--- program plaizgr (robot Fanuc LR Mate 200iD/7L) ---
  Suave(1)
  Establecer velocidad (1000.0 mm/s)
  Est. Ref.: RobotiQ 2F-140 Gripper (Mechanism) Base
  Est. herr: Tool 1
  Mostrar Tool 1
  MoveJ 1 to (362.78, 154.32, 254.42) mm, rotated rx 150.39 ry -54.39 rz -78.94 deg; joints [58.46, 52.97, -15.965, -58.774, -88.343, 127.064]
  MoveL 2 to (362.78, 154.32, 254.42) mm, rotated rx 150.39 ry -54.39 rz -78.94 deg; joints [58.46, 52.97, -15.965, -58.774, -88.343, 127.064]
  MoveL 3 to (343.17, 154.32, 156.36) mm, rotated rx 150.39 ry -54.39 rz -78.94 deg; joints [59.167, 60.189, -23.258, -59.407, -84.021, 132.99]
  MoveL 4 to (343.17, 154.32, 156.36) mm, rotated rx 150.39 ry -54.39 rz -78.94 deg; joints [59.167, 60.189, -23.258, -59.407, -84.021, 132.99]
  Establecer velocidad (50.0 mm/s)
  MoveL 5 to (357.24, 155.51, 156.36) mm, rotated rx 150.39 ry -54.39 rz -78.94 deg; joints [58.593, 58.357, -25.001, -59.364, -83.585, 134.768]
  MoveL 6 to (371.41, 155.49, 156.36) mm, rotated rx 150.39 ry -54.39 rz -78.94 deg; joints [58.07, 56.537, -26.718, -59.336, -83.115, 136.496]
  MoveL 7 to (385.52, 154.28, 156.36) mm, rotated rx 150.39 ry -54.39 rz -78.94 deg; joints [57.607, 54.737, -28.4, -59.33, -82.61, 138.165]
  MoveL 8 to (399.43, 151.88, 156.36) mm, rotated rx 150.39 ry -54.39 rz -78.94 deg; joints [57.21, 52.967, -30.039, -59.349, -82.072, 139.766]
  MoveL 9 to (413.04, 148.32, 157.01) mm, rotated rx 150.39 ry -54.39 rz -78.94 deg; joints [56.883, 51.186, -31.573, -59.393, -81.532, 141.244]
  MoveL 10 to (427.09, 143.6, 159.01) mm, rotated rx 150.39 ry -54.39 rz -78.94 deg; joints [56.601, 49.261, -33.008, -59.45, -81.007, 142.617]
  MoveL 11 to (441.01, 139.44, 162.37) mm, rotated rx 150.39 ry -54.39 rz -78.94 deg; joints [56.277, 47.356, -34.183, -59.457, -80.642, 143.78]
  MoveL 12 to (454.79, 136.05, 167.07) mm, rotated rx 150.39 ry -54.39 rz -78.94 deg; joints [55.897, 45.467, -35.092, -59.397, -80.449, 144.736]
  MoveL 13 to (468.79, 133.33, 171.26) mm, rotated rx 150.39 ry -54.39 rz -78.94 deg; joints [55.448, 43.671, -35.961, -59.295, -80.321, 145.682]
  MoveL 14 to (483.13, 131.27, 174.06) mm, rotated rx 150.39 ry -54.39 rz -78.94 deg; joints [54.922, 42.013, -36.897, -59.158, -80.205, 146.718]
  MoveL 15 to (497.82, 129.91, 175.45) mm, rotated rx 150.39 ry -54.39 rz -78.94 deg; joints [54.312, 40.498, -37.91, -58.981, -80.1, 147.853]
  MoveL 16 to (513.8, 129.29, 175.6) mm, rotated rx 150.39 ry -54.39 rz -78.94 deg; joints [53.565, 39.04, -39.056, -58.741, -80.008, 149.156]
  MoveL 17 to (529.8, 129.54, 175.6) mm, rotated rx 150.39 ry -54.39 rz -78.94 deg; joints [52.727, 37.685, -40.126, -58.427, -80.002, 150.425]
  MoveL 18 to (545.79, 129.54, 175.6) mm, rotated rx 150.39 ry -54.39 rz -78.94 deg; joints [51.873, 36.349, -41.162, -58.086, -80.008, 151.666]
  MoveL 19 to (561.78, 129.54, 175.6) mm, rotated rx 150.39 ry -54.39 rz -78.94 deg; joints [50.985, 35.046, -42.154, -57.706, -80.042, 152.877]
  MoveL 20 to (577.78, 129.54, 175.6) mm, rotated rx 150.39 ry -54.39 rz -78.94 deg; joints [50.063, 33.774, -43.105, -57.286, -80.104, 154.061]
  MoveL 21 to (587.78, 129.54, 175.6) mm, rotated rx 150.39 ry -54.39 rz -78.94 deg; joints [49.468, 32.995, -43.678, -57.001, -80.156, 154.788]
  MoveL 22 to (597.77, 129.54, 175.6) mm, rotated rx 150.39 ry -54.39 rz -78.94 deg; joints [48.857, 32.226, -44.236, -56.7, -80.219, 155.506]
  MoveL 23 to (607.77, 129.54, 175.6) mm, rotated rx 150.39 ry -54.39 rz -78.94 deg; joints [48.232, 31.469, -44.779, -56.382, -80.292, 156.215]
  MoveL 24 to (617.86, 129.25, 175.6) mm, rotated rx 150.39 ry -54.39 rz -78.94 deg; joints [47.606, 30.696, -45.325, -56.058, -80.356, 156.925]
  MoveL 25 to (624.85, 127.52, 175.6) mm, rotated rx 150.39 ry -54.39 rz -78.94 deg; joints [47.271, 30.062, -45.767, -55.904, -80.303, 157.429]
  MoveL 26 to (631.59, 124.12, 175.6) mm, rotated rx 150.39 ry -54.39 rz -78.94 deg; joints [47.066, 29.337, -46.266, -55.841, -80.141, 157.929]
  MoveL 27 to (637.51, 119.15, 175.6) mm, rotated rx 150.39 ry -54.39 rz -78.94 deg; joints [47.027, 28.568, -46.786, -55.891, -79.871, 158.382]
  MoveL 28 to (642.09, 112.97, 175.6) mm, rotated rx 150.39 ry -54.39 rz -78.94 deg; joints [47.169, 27.817, -47.287, -56.061, -79.51, 158.749]
  MoveL 29 to (645.05, 106.13, 175.6) mm, rotated rx 150.39 ry -54.39 rz -78.94 deg; joints [47.477, 27.141, -47.73, -56.336, -79.091, 159.006]
  MoveL 30 to (646.36, 99.2, 175.6) mm, rotated rx 150.39 ry -54.39 rz -78.94 deg; joints [47.914, 26.584, -48.09, -56.687, -78.648, 159.147]
  MoveL 31 to (646.47, 92.51, 175.6) mm, rotated rx 150.39 ry -54.39 rz -78.94 deg; joints [48.424, 26.135, -48.377, -57.079, -78.207, 159.203]
  MoveL 32 to (646.47, 85.85, 175.6) mm, rotated rx 150.39 ry -54.39 rz -78.94 deg; joints [48.949, 25.7, -48.651, -57.481, -77.766, 159.247]
  MoveL 33 to (645.82, 79.04, 175.6) mm, rotated rx 150.39 ry -54.39 rz -78.94 deg; joints [49.539, 25.31, -48.895, -57.924, -77.307, 159.245]
  MoveL 34 to (643.6, 72.09, 175.6) mm, rotated rx 150.39 ry -54.39 rz -78.94 deg; joints [50.256, 25.036, -49.065, -58.442, -76.818, 159.139]
  MoveL 35 to (639.71, 65.55, 175.6) mm, rotated rx 150.39 ry -54.39 rz -78.94 deg; joints [51.058, 24.923, -49.134, -58.997, -76.332, 158.919]
  MoveL 36 to (634.33, 59.99, 175.6) mm, rotated rx 150.39 ry -54.39 rz -78.94 deg; joints [51.88, 24.997, -49.089, -59.541, -75.893, 158.595]
  MoveL 37 to (627.87, 55.87, 175.6) mm, rotated rx 150.39 ry -54.39 rz -78.94 deg; joints [52.646, 25.253, -48.931, -60.02, -75.539, 158.193]
  MoveL 38 to (620.92, 53.42, 175.6) mm, rotated rx 150.39 ry -54.39 rz -78.94 deg; joints [53.296, 25.655, -48.679, -60.397, -75.292, 157.748]
  MoveL 39 to (611.8, 52.57, 175.6) mm, rotated rx 150.39 ry -54.39 rz -78.94 deg; joints [53.933, 26.331, -48.252, -60.721, -75.134, 157.149]
  MoveL 40 to (602.92, 52.57, 175.6) mm, rotated rx 150.39 ry -54.39 rz -78.94 deg; joints [54.47, 27.044, -47.793, -60.966, -75.045, 156.553]
  MoveL 41 to (594.03, 52.57, 175.6) mm, rotated rx 150.39 ry -54.39 rz -78.94 deg; joints [54.993, 27.763, -47.322, -61.196, -74.963, 155.949]
  MoveL 42 to (585.15, 52.57, 175.6) mm, rotated rx 150.39 ry -54.39 rz -78.94 deg; joints [55.503, 28.488, -46.839, -61.411, -74.89, 155.338]
  MoveL 43 to (576.26, 52.57, 175.6) mm, rotated rx 150.39 ry -54.39 rz -78.94 deg; joints [56, 29.22, -46.345, -61.61, -74.826, 154.719]
  MoveL 44 to (567.37, 52.57, 175.6) mm, rotated rx 150.39 ry -54.39 rz -78.94 deg; joints [56.485, 29.958, -45.838, -61.795, -74.77, 154.092]
  MoveL 45 to (549.78, 52.57, 175.6) mm, rotated rx 150.39 ry -54.39 rz -78.94 deg; joints [57.409, 31.439, -44.799, -62.118, -74.685, 152.825]
  MoveL 46 to (532.19, 52.57, 175.6) mm, rotated rx 150.39 ry -54.39 rz -78.94 deg; joints [58.288, 32.948, -43.711, -62.387, -74.634, 151.522]
  MoveL 47 to (514.6, 51.98, 175.6) mm, rotated rx 150.39 ry -54.39 rz -78.94 deg; joints [59.172, 34.456, -42.597, -62.638, -74.577, 150.188]
  MoveL 48 to (497.1, 50.19, 175.42) mm, rotated rx 150.39 ry -54.39 rz -78.94 deg; joints [60.103, 35.943, -41.504, -62.905, -74.462, 148.851]
  MoveL 49 to (482.53, 47.78, 173.97) mm, rotated rx 150.39 ry -54.39 rz -78.94 deg; joints [60.918, 37.26, -40.73, -63.17, -74.265, 147.846]
  MoveL 50 to (468.32, 44.58, 171.14) mm, rotated rx 150.39 ry -54.39 rz -78.94 deg; joints [61.75, 38.633, -40.118, -63.472, -73.975, 146.983]
  MoveL 51 to (454.47, 40.81, 166.96) mm, rotated rx 150.39 ry -54.39 rz -78.94 deg; joints [62.583, 40.068, -39.653, -63.803, -73.608, 146.252]
  MoveL 52 to (440.68, 37.6, 162.27) mm, rotated rx 150.39 ry -54.39 rz -78.94 deg; joints [63.348, 41.583, -39.17, -64.082, -73.29, 145.529]
  MoveL 53 to (426.53, 35.07, 158.91) mm, rotated rx 150.39 ry -54.39 rz -78.94 deg; joints [64.051, 43.092, -38.442, -64.253, -73.114, 144.595]
  MoveL 54 to (412.03, 33.26, 156.92) mm, rotated rx 150.39 ry -54.39 rz -78.94 deg; joints [64.691, 44.6, -37.461, -64.312, -73.085, 143.443]
  MoveL 55 to (398.77, 32.28, 156.36) mm, rotated rx 150.39 ry -54.39 rz -78.94 deg; joints [65.208, 45.953, -36.366, -64.269, -73.187, 142.224]
  MoveL 56 to (385.41, 31.95, 156.36) mm, rotated rx 150.39 ry -54.39 rz -78.94 deg; joints [65.666, 47.346, -35.133, -64.155, -73.389, 140.896]
  MoveL 57 to (372.04, 31.95, 156.36) mm, rotated rx 150.39 ry -54.39 rz -78.94 deg; joints [66.087, 48.8, -33.833, -64.002, -73.645, 139.518]
  MoveL 58 to (358.69, 32.67, 156.36) mm, rotated rx 150.39 ry -54.39 rz -78.94 deg; joints [66.445, 50.337, -32.444, -63.797, -73.987, 138.083]
  MoveL 59 to (345.52, 34.92, 156.36) mm, rotated rx 150.39 ry -54.39 rz -78.94 deg; joints [66.681, 51.991, -30.936, -63.515, -74.476, 136.586]
  MoveL 60 to (332.7, 38.67, 156.6) mm, rotated rx 150.39 ry -54.39 rz -78.94 deg; joints [66.799, 53.734, -29.294, -63.163, -75.121, 135.017]
  MoveL 61 to (320.47, 43.84, 157.41) mm, rotated rx 150.39 ry -54.39 rz -78.94 deg; joints [66.804, 55.532, -27.502, -62.753, -75.932, 133.367]
  MoveL 62 to (308.86, 50.4, 158.71) mm, rotated rx 150.39 ry -54.39 rz -78.94 deg; joints [66.702, 57.406, -25.557, -62.3, -76.911, 131.635]
  MoveL 63 to (298.17, 58.18, 160.36) mm, rotated rx 150.39 ry -54.39 rz -78.94 deg; joints [66.5, 59.336, -23.495, -61.831, -78.04, 129.858]
  MoveL 64 to (292.24, 63.38, 161.47) mm, rotated rx 150.39 ry -54.39 rz -78.94 deg; joints [66.334, 60.525, -22.206, -61.549, -78.785, 128.773]
  MoveL 65 to (286.67, 68.99, 162.65) mm, rotated rx 150.39 ry -54.39 rz -78.94 deg; joints [66.137, 61.748, -20.872, -61.269, -79.585, 127.67]
  MoveL 66 to (281.5, 75.04, 163.85) mm, rotated rx 150.39 ry -54.39 rz -78.94 deg; joints [65.905, 63.007, -19.494, -60.995, -80.441, 126.552]
  MoveL 67 to (277.65, 82.01, 164.81) mm, rotated rx 150.39 ry -54.39 rz -78.94 deg; joints [65.584, 64.2, -18.21, -60.735, -81.331, 125.565]
  MoveL 68 to (275.64, 89.74, 165.34) mm, rotated rx 150.39 ry -54.39 rz -78.94 deg; joints [65.171, 65.21, -17.158, -60.505, -82.19, 124.834]
  MoveL 69 to (275.38, 98.68, 165.41) mm, rotated rx 150.39 ry -54.39 rz -78.94 deg; joints [64.641, 66.072, -16.31, -60.289, -83.05, 124.343]
  MoveL 70 to (276.08, 107.58, 165.22) mm, rotated rx 150.39 ry -54.39 rz -78.94 deg; joints [64.09, 66.803, -15.623, -60.1, -83.851, 124.009]
  MoveL 71 to (278.34, 116.18, 164.63) mm, rotated rx 150.39 ry -54.39 rz -78.94 deg; joints [63.516, 67.235, -15.282, -59.945, -84.501, 123.989]
  MoveL 72 to (282.07, 124.17, 163.71) mm, rotated rx 150.39 ry -54.39 rz -78.94 deg; joints [62.935, 67.338, -15.309, -59.82, -84.972, 124.295]
  MoveL 73 to (287.15, 131.38, 162.54) mm, rotated rx 150.39 ry -54.39 rz -78.94 deg; joints [62.36, 67.11, -15.694, -59.718, -85.258, 124.909]
  MoveL 74 to (293.41, 137.55, 161.24) mm, rotated rx 150.39 ry -54.39 rz -78.94 deg; joints [61.806, 66.572, -16.4, -59.637, -85.36, 125.79]
  MoveL 75 to (300.66, 142.52, 159.94) mm, rotated rx 150.39 ry -54.39 rz -78.94 deg; joints [61.288, 65.764, -17.371, -59.576, -85.297, 126.882]
  MoveL 76 to (308.69, 146.14, 158.73) mm, rotated rx 150.39 ry -54.39 rz -78.94 deg; joints [60.818, 64.735, -18.541, -59.535, -85.089, 128.122]
  MoveL 77 to (317.12, 148.87, 157.73) mm, rotated rx 150.39 ry -54.39 rz -78.94 deg; joints [60.381, 63.612, -19.772, -59.503, -84.821, 129.397]
  MoveL 78 to (325.68, 151.14, 157) mm, rotated rx 150.39 ry -54.39 rz -78.94 deg; joints [59.96, 62.482, -20.966, -59.471, -84.554, 130.631]
  MoveL 79 to (334.36, 152.96, 156.54) mm, rotated rx 150.39 ry -54.39 rz -78.94 deg; joints [59.556, 61.343, -22.128, -59.439, -84.288, 131.829]
  MoveL 80 to (343.17, 154.32, 156.36) mm, rotated rx 150.39 ry -54.39 rz -78.94 deg; joints [59.167, 60.189, -23.258, -59.407, -84.021, 132.99]
  Establecer velocidad (1000.0 mm/s)
  MoveL 81 to (343.17, 154.32, 156.36) mm, rotated rx 150.39 ry -54.39 rz -78.94 deg; joints [59.167, 60.189, -23.258, -59.407, -84.021, 132.99]
  MoveL 82 to (362.78, 154.32, 254.42) mm, rotated rx 150.39 ry -54.39 rz -78.94 deg; joints [58.46, 52.97, -15.965, -58.774, -88.343, 127.064]
  Establecer velocidad (1000.0 mm/s)
  MoveL 83 to (592.37, 52.35, 332.76) mm, rotated rx 150.39 ry -54.39 rz -78.94 deg; joints [55.107, 16.736, -27.061, -58.167, -85.196, 138.168]
  MoveL 84 to (572.75, 52.35, 234.7) mm, rotated rx 150.39 ry -54.39 rz -78.94 deg; joints [56.211, 24.703, -38.872, -60.175, -78.33, 147.93]
  MoveL 85 to (572.75, 52.35, 234.7) mm, rotated rx 150.39 ry -54.39 rz -78.94 deg; joints [56.211, 24.703, -38.872, -60.175, -78.33, 147.93]
  Establecer velocidad (50.0 mm/s)
  MoveL 86 to (566.41, 52.35, 234.7) mm, rotated rx 150.39 ry -54.39 rz -78.94 deg; joints [56.554, 25.28, -38.565, -60.307, -78.25, 147.522]
  MoveL 87 to (560.62, 52.35, 234.7) mm, rotated rx 150.39 ry -54.39 rz -78.94 deg; joints [56.862, 25.81, -38.278, -60.421, -78.182, 147.146]
  MoveL 88 to (556.01, 52.35, 234.7) mm, rotated rx 150.39 ry -54.39 rz -78.94 deg; joints [57.104, 26.234, -38.046, -60.509, -78.131, 146.843]
  MoveL 89 to (552.42, 52.35, 234.7) mm, rotated rx 150.39 ry -54.39 rz -78.94 deg; joints [57.291, 26.566, -37.862, -60.574, -78.093, 146.605]
  MoveL 90 to (548.28, 52.38, 234.7) mm, rotated rx 150.39 ry -54.39 rz -78.94 deg; joints [57.5, 26.951, -37.646, -60.646, -78.055, 146.33]
  MoveL 91 to (543.85, 52.63, 234.7) mm, rotated rx 150.39 ry -54.39 rz -78.94 deg; joints [57.705, 27.377, -37.404, -60.709, -78.032, 146.034]
  MoveL 92 to (538.19, 53.36, 234.7) mm, rotated rx 150.39 ry -54.39 rz -78.94 deg; joints [57.93, 27.948, -37.076, -60.766, -78.036, 145.651]
  MoveL 93 to (531.07, 54.97, 234.7) mm, rotated rx 150.39 ry -54.39 rz -78.94 deg; joints [58.154, 28.71, -36.631, -60.8, -78.097, 145.165]
  MoveL 94 to (524.58, 56.54, 234.7) mm, rotated rx 150.39 ry -54.39 rz -78.94 deg; joints [58.345, 29.413, -36.212, -60.82, -78.167, 144.714]
  MoveL 95 to (518.16, 57.77, 234.7) mm, rotated rx 150.39 ry -54.39 rz -78.94 deg; joints [58.555, 30.095, -35.799, -60.851, -78.22, 144.261]
  MoveL 96 to (511.62, 57.63, 234.7) mm, rotated rx 150.39 ry -54.39 rz -78.94 deg; joints [58.873, 30.712, -35.419, -60.941, -78.179, 143.794]
  MoveL 97 to (505.08, 57.42, 234.7) mm, rotated rx 150.39 ry -54.39 rz -78.94 deg; joints [59.19, 31.33, -35.034, -61.027, -78.139, 143.321]
  MoveL 98 to (498.54, 57.2, 234.7) mm, rotated rx 150.39 ry -54.39 rz -78.94 deg; joints [59.503, 31.951, -34.64, -61.107, -78.105, 142.842]
  MoveL 99 to (492, 57.03, 234.7) mm, rotated rx 150.39 ry -54.39 rz -78.94 deg; joints [59.806, 32.581, -34.236, -61.178, -78.08, 142.357]
  MoveL 100 to (486.16, 56.96, 234.7) mm, rotated rx 150.39 ry -54.39 rz -78.94 deg; joints [60.067, 33.152, -33.865, -61.234, -78.07, 141.919]
  MoveL 101 to (480.31, 57.02, 234.7) mm, rotated rx 150.39 ry -54.39 rz -78.94 deg; joints [60.314, 33.736, -33.482, -61.279, -78.074, 141.474]
  MoveL 102 to (474.48, 57.28, 234.7) mm, rotated rx 150.39 ry -54.39 rz -78.94 deg; joints [60.542, 34.334, -33.084, -61.311, -78.098, 141.024]
  MoveL 103 to (468.66, 57.82, 234.7) mm, rotated rx 150.39 ry -54.39 rz -78.94 deg; joints [60.745, 34.95, -32.669, -61.328, -78.147, 140.568]
  MoveL 104 to (462.91, 58.77, 234.7) mm, rotated rx 150.39 ry -54.39 rz -78.94 deg; joints [60.912, 35.589, -32.234, -61.323, -78.232, 140.11]
  MoveL 105 to (457.85, 61.63, 234.7) mm, rotated rx 150.39 ry -54.39 rz -78.94 deg; joints [60.909, 36.269, -31.766, -61.237, -78.46, 139.691]
  MoveL 106 to (454, 66, 234.7) mm, rotated rx 150.39 ry -54.39 rz -78.94 deg; joints [60.747, 36.917, -31.314, -61.086, -78.799, 139.356]
  MoveL 107 to (451.47, 71.25, 234.7) mm, rotated rx 150.39 ry -54.39 rz -78.94 deg; joints [60.472, 37.486, -30.914, -60.898, -79.199, 139.115]
  MoveL 108 to (450.78, 77.03, 234.7) mm, rotated rx 150.39 ry -54.39 rz -78.94 deg; joints [60.088, 37.899, -30.62, -60.684, -79.63, 139.019]
  MoveL 109 to (451.23, 79.92, 234.7) mm, rotated rx 150.39 ry -54.39 rz -78.94 deg; joints [59.864, 38.025, -30.53, -60.573, -79.842, 139.034]
  MoveL 110 to (452.01, 82.76, 234.7) mm, rotated rx 150.39 ry -54.39 rz -78.94 deg; joints [59.632, 38.116, -30.465, -60.462, -80.048, 139.077]
  MoveL 111 to (452.81, 85.6, 234.7) mm, rotated rx 150.39 ry -54.39 rz -78.94 deg; joints [59.399, 38.206, -30.401, -60.352, -80.255, 139.121]
  MoveL 112 to (453.63, 88.43, 234.7) mm, rotated rx 150.39 ry -54.39 rz -78.94 deg; joints [59.166, 38.296, -30.336, -60.242, -80.461, 139.165]
  MoveL 113 to (454.46, 91.26, 234.7) mm, rotated rx 150.39 ry -54.39 rz -78.94 deg; joints [58.933, 38.386, -30.272, -60.132, -80.667, 139.21]
  MoveL 114 to (455.13, 94.08, 234.7) mm, rotated rx 150.39 ry -54.39 rz -78.94 deg; joints [58.709, 38.493, -30.195, -60.024, -80.874, 139.24]
  MoveL 115 to (452.96, 100.35, 234.7) mm, rotated rx 150.39 ry -54.39 rz -78.94 deg; joints [58.367, 39.113, -29.747, -59.815, -81.355, 138.998]
  MoveL 116 to (450.97, 106.68, 234.7) mm, rotated rx 150.39 ry -54.39 rz -78.94 deg; joints [58.019, 39.727, -29.298, -59.609, -81.843, 138.761]
  MoveL 117 to (450.88, 111.09, 234.7) mm, rotated rx 150.39 ry -54.39 rz -78.94 deg; joints [57.724, 40.026, -29.079, -59.457, -82.176, 138.702]
  MoveL 118 to (452.32, 115.26, 234.7) mm, rotated rx 150.39 ry -54.39 rz -78.94 deg; joints [57.381, 40.151, -28.987, -59.3, -82.481, 138.776]
  MoveL 119 to (454.97, 118.8, 234.7) mm, rotated rx 150.39 ry -54.39 rz -78.94 deg; joints [57.029, 40.113, -29.015, -59.153, -82.731, 138.959]
  MoveL 120 to (459.29, 121.86, 234.7) mm, rotated rx 150.39 ry -54.39 rz -78.94 deg; joints [56.635, 39.874, -29.191, -59.003, -82.936, 139.289]
  MoveL 121 to (464.42, 123.12, 234.7) mm, rotated rx 150.39 ry -54.39 rz -78.94 deg; joints [56.323, 39.435, -29.512, -58.902, -83.002, 139.708]
  MoveL 122 to (469.68, 123.65, 234.7) mm, rotated rx 150.39 ry -54.39 rz -78.94 deg; joints [56.052, 38.937, -29.874, -58.82, -83.017, 140.143]
  MoveL 123 to (474.96, 123.96, 234.7) mm, rotated rx 150.39 ry -54.39 rz -78.94 deg; joints [55.791, 38.429, -30.241, -58.742, -83.02, 140.577]
  MoveL 124 to (480.25, 124.12, 234.7) mm, rotated rx 150.39 ry -54.39 rz -78.94 deg; joints [55.537, 37.915, -30.609, -58.666, -83.016, 141.009]
  MoveL 125 to (491.89, 124.14, 234.7) mm, rotated rx 150.39 ry -54.39 rz -78.94 deg; joints [54.989, 36.778, -31.412, -58.497, -82.999, 141.945]
  MoveL 126 to (503.52, 123.96, 234.7) mm, rotated rx 150.39 ry -54.39 rz -78.94 deg; joints [54.439, 35.65, -32.193, -58.32, -82.987, 142.863]
  MoveL 127 to (515.16, 123.84, 234.7) mm, rotated rx 150.39 ry -54.39 rz -78.94 deg; joints [53.87, 34.546, -32.943, -58.123, -83, 143.759]
  MoveL 128 to (526.61, 125.64, 234.7) mm, rotated rx 150.39 ry -54.39 rz -78.94 deg; joints [53.161, 33.611, -33.565, -57.836, -83.173, 144.607]
  MoveL 129 to (538.1, 127.62, 234.7) mm, rotated rx 150.39 ry -54.39 rz -78.94 deg; joints [52.42, 32.703, -34.158, -57.521, -83.376, 145.444]
  MoveL 130 to (549.77, 128.88, 234.7) mm, rotated rx 150.39 ry -54.39 rz -78.94 deg; joints [51.701, 31.748, -34.77, -57.21, -83.545, 146.284]
  MoveL 131 to (569.54, 129.58, 234.7) mm, rotated rx 150.39 ry -54.39 rz -78.94 deg; joints [50.539, 30.071, -35.814, -56.693, -83.771, 147.685]
  MoveL 132 to (589.33, 129.07, 234.7) mm, rotated rx 150.39 ry -54.39 rz -78.94 deg; joints [49.406, 28.352, -36.842, -56.168, -83.963, 149.053]
  MoveL 133 to (597.7, 128.45, 234.7) mm, rotated rx 150.39 ry -54.39 rz -78.94 deg; joints [48.938, 27.608, -37.273, -55.946, -84.032, 149.623]
  MoveL 134 to (606.05, 127.58, 234.7) mm, rotated rx 150.39 ry -54.39 rz -78.94 deg; joints [48.479, 26.854, -37.701, -55.725, -84.093, 150.185]
  MoveL 135 to (614.37, 126.46, 234.7) mm, rotated rx 150.39 ry -54.39 rz -78.94 deg; joints [48.029, 26.09, -38.126, -55.505, -84.146, 150.738]
  MoveL 136 to (622.65, 125.08, 234.7) mm, rotated rx 150.39 ry -54.39 rz -78.94 deg; joints [47.59, 25.317, -38.546, -55.288, -84.191, 151.283]
  MoveL 137 to (630.62, 122.45, 234.7) mm, rotated rx 150.39 ry -54.39 rz -78.94 deg; joints [47.252, 24.48, -38.99, -55.129, -84.154, 151.8]
  MoveL 138 to (637.7, 117.98, 234.7) mm, rotated rx 150.39 ry -54.39 rz -78.94 deg; joints [47.1, 23.582, -39.453, -55.079, -83.986, 152.25]
  MoveL 139 to (642.31, 113.59, 234.7) mm, rotated rx 150.39 ry -54.39 rz -78.94 deg; joints [47.108, 22.887, -39.801, -55.114, -83.782, 152.533]
  MoveL 140 to (646.07, 108.5, 234.7) mm, rotated rx 150.39 ry -54.39 rz -78.94 deg; joints [47.228, 22.209, -40.133, -55.216, -83.517, 152.755]
  MoveL 141 to (648.78, 102.72, 234.7) mm, rotated rx 150.39 ry -54.39 rz -78.94 deg; joints [47.476, 21.565, -40.441, -55.393, -83.185, 152.902]
  MoveL 142 to (650.24, 96.55, 234.7) mm, rotated rx 150.39 ry -54.39 rz -78.94 deg; joints [47.848, 20.994, -40.708, -55.642, -82.802, 152.962]
  MoveL 143 to (650.47, 90.13, 234.7) mm, rotated rx 150.39 ry -54.39 rz -78.94 deg; joints [48.332, 20.507, -40.931, -55.956, -82.374, 152.94]
  MoveL 144 to (649.71, 82.15, 234.7) mm, rotated rx 150.39 ry -54.39 rz -78.94 deg; joints [49.02, 19.994, -41.161, -56.394, -81.815, 152.841]
  MoveL 145 to (646.76, 74.64, 234.7) mm, rotated rx 150.39 ry -54.39 rz -78.94 deg; joints [49.83, 19.706, -41.288, -56.894, -81.236, 152.61]
  MoveL 146 to (641.96, 68.13, 234.7) mm, rotated rx 150.39 ry -54.39 rz -78.94 deg; joints [50.692, 19.654, -41.31, -57.41, -80.679, 152.273]
  MoveL 147 to (635.83, 62.85, 234.7) mm, rotated rx 150.39 ry -54.39 rz -78.94 deg; joints [51.541, 19.814, -41.24, -57.902, -80.178, 151.867]
  MoveL 148 to (628.75, 59.03, 234.7) mm, rotated rx 150.39 ry -54.39 rz -78.94 deg; joints [52.324, 20.165, -41.084, -58.339, -79.76, 151.416]
  MoveL 149 to (620.95, 56.87, 234.7) mm, rotated rx 150.39 ry -54.39 rz -78.94 deg; joints [53.004, 20.699, -40.843, -58.698, -79.448, 150.935]
  MoveL 150 to (596.95, 53.5, 234.7) mm, rotated rx 150.39 ry -54.39 rz -78.94 deg; joints [54.745, 22.598, -39.943, -59.547, -78.771, 149.455]
  MoveL 151 to (572.75, 52.35, 234.7) mm, rotated rx 150.39 ry -54.39 rz -78.94 deg; joints [56.211, 24.703, -38.872, -60.175, -78.33, 147.93]
  Establecer velocidad (1000.0 mm/s)
  MoveL 152 to (572.75, 52.35, 234.7) mm, rotated rx 150.39 ry -54.39 rz -78.94 deg; joints [56.211, 24.703, -38.872, -60.175, -78.33, 147.93]
  MoveL 153 to (592.37, 52.35, 332.76) mm, rotated rx 150.39 ry -54.39 rz -78.94 deg; joints [55.107, 16.736, -27.061, -58.167, -85.196, 138.168]

--- program pladerch (robot Fanuc LR Mate 200iD/7L) ---
  Suave(1)
  Establecer velocidad (1000.0 mm/s)
  Est. Ref.: RobotiQ 2F-140 Gripper (Mechanism) Base
  Est. herr: Tool 1
  Mostrar Tool 1
  MoveJ 1 to (235.91, 212.79, 258.59) mm, rotated rx 164.21 ry -43.9 rz -78.89 deg; joints [57.845, 56.233, -8.401, -42.896, -98.91, 126.65]
  MoveL 2 to (235.91, 212.79, 258.59) mm, rotated rx 164.21 ry -43.9 rz -78.89 deg; joints [57.845, 56.233, -8.401, -42.896, -98.91, 126.65]
  MoveL 3 to (216.3, 212.79, 160.54) mm, rotated rx 164.21 ry -43.9 rz -78.89 deg; joints [58.546, 62.427, -16.246, -42.557, -92.678, 131.492]
  MoveL 4 to (216.3, 212.79, 160.54) mm, rotated rx 164.21 ry -43.9 rz -78.89 deg; joints [58.546, 62.427, -16.246, -42.557, -92.678, 131.492]
  Establecer velocidad (50.0 mm/s)
  MoveL 5 to (225.57, 213.87, 160.54) mm, rotated rx 164.21 ry -43.9 rz -78.89 deg; joints [58.156, 60.991, -17.597, -42.395, -91.933, 132.681]
  MoveL 6 to (234.89, 213.99, 160.54) mm, rotated rx 164.21 ry -43.9 rz -78.89 deg; joints [57.812, 59.541, -18.949, -42.256, -91.154, 133.832]
  MoveL 7 to (244.22, 213.91, 160.54) mm, rotated rx 164.21 ry -43.9 rz -78.89 deg; joints [57.474, 58.154, -20.23, -42.128, -90.418, 134.929]
  MoveL 8 to (253.51, 213.4, 160.69) mm, rotated rx 164.21 ry -43.9 rz -78.89 deg; joints [57.156, 56.795, -21.453, -42.014, -89.71, 135.969]
  MoveL 9 to (263.17, 212.36, 161.72) mm, rotated rx 164.21 ry -43.9 rz -78.89 deg; joints [56.849, 55.36, -22.609, -41.909, -89.041, 136.954]
  MoveL 10 to (272.6, 210.83, 163.66) mm, rotated rx 164.21 ry -43.9 rz -78.89 deg; joints [56.573, 53.925, -23.618, -41.82, -88.459, 137.816]
  MoveL 11 to (281.78, 208.84, 166.52) mm, rotated rx 164.21 ry -43.9 rz -78.89 deg; joints [56.328, 52.48, -24.486, -41.743, -87.96, 138.561]
  MoveL 12 to (290.87, 206.4, 169.55) mm, rotated rx 164.21 ry -43.9 rz -78.89 deg; joints [56.109, 51.041, -25.304, -41.679, -87.481, 139.255]
  MoveL 13 to (300.19, 204.13, 171.69) mm, rotated rx 164.21 ry -43.9 rz -78.89 deg; joints [55.865, 49.671, -26.171, -41.608, -86.98, 139.996]
  MoveL 14 to (309.75, 202.38, 172.93) mm, rotated rx 164.21 ry -43.9 rz -78.89 deg; joints [55.574, 48.397, -27.073, -41.523, -86.478, 140.79]
  MoveL 15 to (320.22, 201.09, 173.24) mm, rotated rx 164.21 ry -43.9 rz -78.89 deg; joints [55.207, 47.142, -28.08, -41.414, -85.938, 141.703]
  MoveL 16 to (330.77, 200.46, 173.24) mm, rotated rx 164.21 ry -43.9 rz -78.89 deg; joints [54.788, 45.978, -29.044, -41.282, -85.458, 142.619]
  MoveL 17 to (341.34, 200.38, 173.24) mm, rotated rx 164.21 ry -43.9 rz -78.89 deg; joints [54.322, 44.884, -29.94, -41.127, -85.051, 143.517]
  MoveL 18 to (351.91, 200.38, 173.24) mm, rotated rx 164.21 ry -43.9 rz -78.89 deg; joints [53.84, 43.822, -30.799, -40.962, -84.676, 144.398]
  MoveL 19 to (362.48, 200.38, 173.24) mm, rotated rx 164.21 ry -43.9 rz -78.89 deg; joints [53.348, 42.786, -31.628, -40.79, -84.325, 145.263]
  MoveL 20 to (388.9, 200.38, 173.24) mm, rotated rx 164.21 ry -43.9 rz -78.89 deg; joints [52.064, 40.294, -33.579, -40.32, -83.546, 147.365]
  MoveL 21 to (393.41, 200.03, 173.24) mm, rotated rx 164.21 ry -43.9 rz -78.89 deg; joints [51.86, 39.856, -33.915, -40.247, -83.399, 147.714]
  MoveL 22 to (398.02, 198.64, 173.24) mm, rotated rx 164.21 ry -43.9 rz -78.89 deg; joints [51.715, 39.339, -34.31, -40.206, -83.175, 148.063]
  MoveL 23 to (402.39, 196.15, 173.24) mm, rotated rx 164.21 ry -43.9 rz -78.89 deg; joints [51.653, 38.769, -34.741, -40.21, -82.878, 148.383]
  MoveL 24 to (406.12, 192.66, 173.24) mm, rotated rx 164.21 ry -43.9 rz -78.89 deg; joints [51.688, 38.19, -35.177, -40.263, -82.527, 148.645]
  MoveL 25 to (408.92, 188.44, 173.24) mm, rotated rx 164.21 ry -43.9 rz -78.89 deg; joints [51.821, 37.647, -35.582, -40.364, -82.149, 148.825]
  MoveL 26 to (410.62, 183.87, 173.24) mm, rotated rx 164.21 ry -43.9 rz -78.89 deg; joints [52.037, 37.18, -35.927, -40.503, -81.773, 148.917]
  MoveL 27 to (411.25, 179.33, 173.24) mm, rotated rx 164.21 ry -43.9 rz -78.89 deg; joints [52.308, 36.813, -36.197, -40.664, -81.425, 148.926]
  MoveL 28 to (411.26, 174.92, 173.24) mm, rotated rx 164.21 ry -43.9 rz -78.89 deg; joints [52.605, 36.513, -36.416, -40.834, -81.102, 148.887]
  MoveL 29 to (411.24, 170.52, 173.24) mm, rotated rx 164.21 ry -43.9 rz -78.89 deg; joints [52.907, 36.218, -36.631, -41.007, -80.781, 148.844]
  MoveL 30 to (410.58, 165.97, 173.24) mm, rotated rx 164.21 ry -43.9 rz -78.89 deg; joints [53.253, 35.974, -36.808, -41.199, -80.466, 148.75]
  MoveL 31 to (408.85, 161.41, 173.24) mm, rotated rx 164.21 ry -43.9 rz -78.89 deg; joints [53.658, 35.827, -36.914, -41.412, -80.172, 148.575]
  MoveL 32 to (406.03, 157.2, 173.24) mm, rotated rx 164.21 ry -43.9 rz -78.89 deg; joints [54.094, 35.805, -36.929, -41.63, -79.929, 148.32]
  MoveL 33 to (402.28, 153.74, 173.24) mm, rotated rx 164.21 ry -43.9 rz -78.89 deg; joints [54.526, 35.919, -36.847, -41.833, -79.761, 148.003]
  MoveL 34 to (397.9, 151.27, 173.24) mm, rotated rx 164.21 ry -43.9 rz -78.89 deg; joints [54.916, 36.157, -36.675, -42.004, -79.68, 147.649]
  MoveL 35 to (392.62, 149.81, 173.24) mm, rotated rx 164.21 ry -43.9 rz -78.89 deg; joints [55.277, 36.545, -36.393, -42.145, -79.695, 147.238]
  MoveL 36 to (387.52, 149.58, 173.24) mm, rotated rx 164.21 ry -43.9 rz -78.89 deg; joints [55.54, 36.999, -36.06, -42.231, -79.799, 146.851]
  MoveL 37 to (382.49, 149.58, 173.24) mm, rotated rx 164.21 ry -43.9 rz -78.89 deg; joints [55.78, 37.465, -35.716, -42.305, -79.923, 146.47]
  MoveL 38 to (377.46, 149.58, 173.24) mm, rotated rx 164.21 ry -43.9 rz -78.89 deg; joints [56.017, 37.935, -35.367, -42.376, -80.051, 146.087]
  MoveL 39 to (372.42, 149.58, 173.24) mm, rotated rx 164.21 ry -43.9 rz -78.89 deg; joints [56.252, 38.408, -35.013, -42.445, -80.183, 145.7]
  MoveL 40 to (367.39, 149.58, 173.24) mm, rotated rx 164.21 ry -43.9 rz -78.89 deg; joints [56.483, 38.886, -34.653, -42.511, -80.32, 145.312]
  MoveL 41 to (362.36, 149.58, 173.24) mm, rotated rx 164.21 ry -43.9 rz -78.89 deg; joints [56.712, 39.368, -34.287, -42.576, -80.462, 144.92]
  MoveL 42 to (350.73, 149.58, 173.24) mm, rotated rx 164.21 ry -43.9 rz -78.89 deg; joints [57.23, 40.497, -33.421, -42.715, -80.808, 144.005]
  MoveL 43 to (339.1, 149.58, 173.24) mm, rotated rx 164.21 ry -43.9 rz -78.89 deg; joints [57.734, 41.652, -32.523, -42.844, -81.18, 143.073]
  MoveL 44 to (327.48, 149.75, 173.24) mm, rotated rx 164.21 ry -43.9 rz -78.89 deg; joints [58.213, 42.843, -31.582, -42.956, -81.593, 142.124]
  MoveL 45 to (315.86, 149.49, 173.22) mm, rotated rx 164.21 ry -43.9 rz -78.89 deg; joints [58.707, 44.037, -30.628, -43.072, -82.002, 141.154]
  MoveL 46 to (306.09, 148.73, 172.57) mm, rotated rx 164.21 ry -43.9 rz -78.89 deg; joints [59.148, 45.068, -29.89, -43.187, -82.28, 140.364]
  MoveL 47 to (296.55, 147.49, 170.97) mm, rotated rx 164.21 ry -43.9 rz -78.89 deg; joints [59.603, 46.119, -29.265, -43.315, -82.464, 139.642]
  MoveL 48 to (287.24, 145.81, 168.45) mm, rotated rx 164.21 ry -43.9 rz -78.89 deg; joints [60.068, 47.19, -28.749, -43.456, -82.56, 138.985]
  MoveL 49 to (278.12, 143.7, 165.26) mm, rotated rx 164.21 ry -43.9 rz -78.89 deg; joints [60.546, 48.27, -28.311, -43.605, -82.588, 138.374]
  MoveL 50 to (268.95, 141.09, 162.8) mm, rotated rx 164.21 ry -43.9 rz -78.89 deg; joints [61.05, 49.303, -27.793, -43.754, -82.656, 137.689]
  MoveL 51 to (259.7, 137.99, 161.24) mm, rotated rx 164.21 ry -43.9 rz -78.89 deg; joints [61.579, 50.285, -27.174, -43.9, -82.777, 136.916]
  MoveL 52 to (249.54, 135.14, 160.55) mm, rotated rx 164.21 ry -43.9 rz -78.89 deg; joints [62.115, 51.373, -26.326, -44.025, -83.056, 135.975]
  MoveL 53 to (239.11, 133.26, 160.54) mm, rotated rx 164.21 ry -43.9 rz -78.89 deg; joints [62.586, 52.559, -25.282, -44.109, -83.511, 134.938]
  MoveL 54 to (228.51, 132.4, 160.54) mm, rotated rx 164.21 ry -43.9 rz -78.89 deg; joints [62.988, 53.882, -24.105, -44.16, -84.1, 133.849]
  MoveL 55 to (217.88, 132.57, 160.54) mm, rotated rx 164.21 ry -43.9 rz -78.89 deg; joints [63.318, 55.339, -22.797, -44.181, -84.828, 132.715]
  MoveL 56 to (207.36, 133.76, 160.59) mm, rotated rx 164.21 ry -43.9 rz -78.89 deg; joints [63.573, 56.922, -21.351, -44.18, -85.7, 131.534]
  MoveL 57 to (200.91, 135, 160.87) mm, rotated rx 164.21 ry -43.9 rz -78.89 deg; joints [63.695, 57.965, -20.357, -44.169, -86.334, 130.758]
  MoveL 58 to (194.56, 136.62, 161.37) mm, rotated rx 164.21 ry -43.9 rz -78.89 deg; joints [63.788, 59.051, -19.284, -44.154, -87.042, 129.947]
  MoveL 59 to (188.32, 138.61, 162.1) mm, rotated rx 164.21 ry -43.9 rz -78.89 deg; joints [63.854, 60.192, -18.124, -44.137, -87.831, 129.093]
  MoveL 60 to (182.41, 141.35, 163) mm, rotated rx 164.21 ry -43.9 rz -78.89 deg; joints [63.864, 61.389, -16.881, -44.113, -88.718, 128.22]
  MoveL 61 to (177.16, 145.2, 163.97) mm, rotated rx 164.21 ry -43.9 rz -78.89 deg; joints [63.787, 62.638, -15.571, -44.08, -89.709, 127.362]
  MoveL 62 to (172.79, 149.99, 164.9) mm, rotated rx 164.21 ry -43.9 rz -78.89 deg; joints [63.629, 63.892, -14.254, -44.043, -90.762, 126.555]
  MoveL 63 to (169.43, 155.61, 165.7) mm, rotated rx 164.21 ry -43.9 rz -78.89 deg; joints [63.395, 65.121, -12.972, -44.004, -91.842, 125.828]
  MoveL 64 to (167.25, 161.76, 166.26) mm, rotated rx 164.21 ry -43.9 rz -78.89 deg; joints [63.097, 66.253, -11.81, -43.965, -92.88, 125.229]
  MoveL 65 to (166.5, 166.11, 166.46) mm, rotated rx 164.21 ry -43.9 rz -78.89 deg; joints [62.866, 66.929, -11.13, -43.936, -93.527, 124.921]
  MoveL 66 to (166.32, 170.52, 166.51) mm, rotated rx 164.21 ry -43.9 rz -78.89 deg; joints [62.614, 67.512, -10.559, -43.904, -94.11, 124.702]
  MoveL 67 to (166.39, 174.93, 166.49) mm, rotated rx 164.21 ry -43.9 rz -78.89 deg; joints [62.356, 68.063, -10.027, -43.872, -94.669, 124.516]
  MoveL 68 to (167.21, 179.23, 166.27) mm, rotated rx 164.21 ry -43.9 rz -78.89 deg; joints [62.083, 68.435, -9.694, -43.828, -95.095, 124.479]
  MoveL 69 to (169.65, 184.52, 165.65) mm, rotated rx 164.21 ry -43.9 rz -78.89 deg; joints [61.704, 68.55, -9.667, -43.741, -95.374, 124.731]
  MoveL 70 to (173.3, 189.04, 164.79) mm, rotated rx 164.21 ry -43.9 rz -78.89 deg; joints [61.332, 68.267, -10.061, -43.627, -95.342, 125.27]
  MoveL 71 to (177.35, 193.16, 163.93) mm, rotated rx 164.21 ry -43.9 rz -78.89 deg; joints [60.968, 67.852, -10.582, -43.505, -95.211, 125.891]
  MoveL 72 to (183.97, 198.73, 162.74) mm, rotated rx 164.21 ry -43.9 rz -78.89 deg; joints [60.439, 67.068, -11.505, -43.314, -94.898, 126.907]
  MoveL 73 to (191.25, 203.56, 161.73) mm, rotated rx 164.21 ry -43.9 rz -78.89 deg; joints [59.925, 66.109, -12.57, -43.117, -94.466, 128.006]
  MoveL 74 to (199.05, 207.53, 160.99) mm, rotated rx 164.21 ry -43.9 rz -78.89 deg; joints [59.439, 65.012, -13.725, -42.923, -93.944, 129.143]
  MoveL 75 to (207.24, 210.58, 160.59) mm, rotated rx 164.21 ry -43.9 rz -78.89 deg; joints [58.986, 63.806, -14.931, -42.738, -93.358, 130.287]
  Establecer velocidad (1000.0 mm/s)
  MoveL 76 to (207.24, 210.58, 160.59) mm, rotated rx 164.21 ry -43.9 rz -78.89 deg; joints [58.986, 63.806, -14.931, -42.738, -93.358, 130.287]
  MoveL 77 to (226.85, 210.58, 258.65) mm, rotated rx 164.21 ry -43.9 rz -78.89 deg; joints [58.299, 57.675, -7.13, -43.152, -99.532, 125.438]
  Establecer velocidad (1000.0 mm/s)
  MoveL 78 to (382.21, 200.52, 310.42) mm, rotated rx 164.21 ry -43.9 rz -78.89 deg; joints [52.387, 34.35, -17.597, -40.379, -95.57, 136.815]
  MoveL 79 to (362.6, 200.52, 212.36) mm, rotated rx 164.21 ry -43.9 rz -78.89 deg; joints [53.333, 40.551, -27.477, -40.589, -87.482, 142.56]
  MoveL 80 to (362.6, 200.52, 212.36) mm, rotated rx 164.21 ry -43.9 rz -78.89 deg; joints [53.333, 40.551, -27.477, -40.589, -87.482, 142.56]
  Establecer velocidad (50.0 mm/s)
  MoveL 81 to (378.48, 199.76, 212.36) mm, rotated rx 164.21 ry -43.9 rz -78.89 deg; joints [52.619, 38.913, -28.667, -40.314, -86.985, 143.813]
  MoveL 82 to (394.24, 197.56, 212.36) mm, rotated rx 164.21 ry -43.9 rz -78.89 deg; joints [51.977, 37.23, -29.858, -40.069, -86.436, 145.011]
  MoveL 83 to (399.36, 196.18, 212.36) mm, rotated rx 164.21 ry -43.9 rz -78.89 deg; joints [51.806, 36.642, -30.265, -40.007, -86.219, 145.388]
  MoveL 84 to (404.03, 193.71, 212.36) mm, rotated rx 164.21 ry -43.9 rz -78.89 deg; joints [51.728, 36.022, -30.691, -39.99, -85.937, 145.714]
  MoveL 85 to (408.09, 190.29, 212.36) mm, rotated rx 164.21 ry -43.9 rz -78.89 deg; joints [51.742, 35.393, -31.118, -40.017, -85.602, 145.979]
  MoveL 86 to (411.28, 186.07, 212.36) mm, rotated rx 164.21 ry -43.9 rz -78.89 deg; joints [51.855, 34.79, -31.523, -40.091, -85.23, 146.167]
  MoveL 87 to (413.3, 181.18, 212.36) mm, rotated rx 164.21 ry -43.9 rz -78.89 deg; joints [52.077, 34.251, -31.88, -40.215, -84.835, 146.254]
  MoveL 88 to (413.89, 175.92, 212.36) mm, rotated rx 164.21 ry -43.9 rz -78.89 deg; joints [52.401, 33.821, -32.163, -40.384, -84.442, 146.226]
  MoveL 89 to (413.64, 170.65, 212.36) mm, rotated rx 164.21 ry -43.9 rz -78.89 deg; joints [52.773, 33.473, -32.39, -40.573, -84.065, 146.134]
  MoveL 90 to (412.13, 165.64, 212.36) mm, rotated rx 164.21 ry -43.9 rz -78.89 deg; joints [53.196, 33.263, -32.526, -40.781, -83.729, 145.951]
  MoveL 91 to (409.35, 161.16, 212.36) mm, rotated rx 164.21 ry -43.9 rz -78.89 deg; joints [53.649, 33.212, -32.559, -40.995, -83.454, 145.682]
  MoveL 92 to (405.67, 157.41, 212.36) mm, rotated rx 164.21 ry -43.9 rz -78.89 deg; joints [54.098, 33.301, -32.501, -41.198, -83.249, 145.357]
  MoveL 93 to (401.4, 154.59, 212.36) mm, rotated rx 164.21 ry -43.9 rz -78.89 deg; joints [54.51, 33.512, -32.364, -41.377, -83.122, 145.003]
  MoveL 94 to (396.62, 152.78, 212.36) mm, rotated rx 164.21 ry -43.9 rz -78.89 deg; joints [54.873, 33.844, -32.148, -41.526, -83.081, 144.626]
  MoveL 95 to (391.62, 151.87, 212.36) mm, rotated rx 164.21 ry -43.9 rz -78.89 deg; joints [55.181, 34.26, -31.874, -41.644, -83.113, 144.246]
  MoveL 96 to (386.59, 151.14, 212.36) mm, rotated rx 164.21 ry -43.9 rz -78.89 deg; joints [55.475, 34.696, -31.585, -41.753, -83.162, 143.865]
  MoveL 97 to (373.7, 149.91, 212.36) mm, rotated rx 164.21 ry -43.9 rz -78.89 deg; joints [56.169, 35.874, -30.792, -41.997, -83.356, 142.887]
  MoveL 98 to (360.76, 149.56, 212.36) mm, rotated rx 164.21 ry -43.9 rz -78.89 deg; joints [56.785, 37.141, -29.919, -42.197, -83.648, 141.901]
  MoveL 99 to (349, 149.91, 212.36) mm, rotated rx 164.21 ry -43.9 rz -78.89 deg; joints [57.283, 38.363, -29.059, -42.345, -83.992, 140.996]
  MoveL 100 to (337.35, 151.21, 212.36) mm, rotated rx 164.21 ry -43.9 rz -78.89 deg; joints [57.699, 39.661, -28.127, -42.453, -84.435, 140.094]
  MoveL 101 to (325.93, 153.37, 212.36) mm, rotated rx 164.21 ry -43.9 rz -78.89 deg; joints [58.035, 41.022, -27.129, -42.526, -84.97, 139.196]
  MoveL 102 to (314.3, 153.24, 212.36) mm, rotated rx 164.21 ry -43.9 rz -78.89 deg; joints [58.521, 42.284, -26.185, -42.663, -85.37, 138.234]
  MoveL 103 to (302.67, 153.18, 212.36) mm, rotated rx 164.21 ry -43.9 rz -78.89 deg; joints [58.99, 43.584, -25.195, -42.79, -85.811, 137.25]
  MoveL 104 to (299.22, 153.26, 212.36) mm, rotated rx 164.21 ry -43.9 rz -78.89 deg; joints [59.12, 43.985, -24.887, -42.824, -85.957, 136.952]
  MoveL 105 to (295.76, 153.43, 212.36) mm, rotated rx 164.21 ry -43.9 rz -78.89 deg; joints [59.243, 44.394, -24.569, -42.855, -86.113, 136.654]
  MoveL 106 to (292.32, 153.73, 212.36) mm, rotated rx 164.21 ry -43.9 rz -78.89 deg; joints [59.357, 44.816, -24.241, -42.882, -86.283, 136.354]
  MoveL 107 to (288.91, 154.29, 212.36) mm, rotated rx 164.21 ry -43.9 rz -78.89 deg; joints [59.452, 45.255, -23.898, -42.902, -86.476, 136.056]
  MoveL 108 to (285.89, 155.93, 212.36) mm, rotated rx 164.21 ry -43.9 rz -78.89 deg; joints [59.461, 45.727, -23.526, -42.89, -86.743, 135.797]
  MoveL 109 to (283.93, 158.04, 212.36) mm, rotated rx 164.21 ry -43.9 rz -78.89 deg; joints [59.4, 46.111, -23.222, -42.857, -87.004, 135.631]
  MoveL 110 to (282.64, 160.61, 212.36) mm, rotated rx 164.21 ry -43.9 rz -78.89 deg; joints [59.284, 46.449, -22.954, -42.806, -87.273, 135.526]
  MoveL 111 to (282.27, 163.45, 212.36) mm, rotated rx 164.21 ry -43.9 rz -78.89 deg; joints [59.116, 46.699, -22.754, -42.74, -87.524, 135.504]
  MoveL 112 to (282.87, 166.27, 212.36) mm, rotated rx 164.21 ry -43.9 rz -78.89 deg; joints [58.914, 46.831, -22.649, -42.665, -87.729, 135.57]
  MoveL 113 to (283.8, 169.02, 212.36) mm, rotated rx 164.21 ry -43.9 rz -78.89 deg; joints [58.704, 46.921, -22.577, -42.588, -87.913, 135.664]
  MoveL 114 to (284.74, 171.76, 212.36) mm, rotated rx 164.21 ry -43.9 rz -78.89 deg; joints [58.494, 47.01, -22.506, -42.51, -88.096, 135.759]
  MoveL 115 to (285, 173.96, 212.36) mm, rotated rx 164.21 ry -43.9 rz -78.89 deg; joints [58.345, 47.142, -22.4, -42.455, -88.267, 135.789]
  MoveL 116 to (284.34, 176.18, 212.36) mm, rotated rx 164.21 ry -43.9 rz -78.89 deg; joints [58.231, 47.389, -22.201, -42.41, -88.485, 135.732]
  MoveL 117 to (283.69, 178.41, 212.36) mm, rotated rx 164.21 ry -43.9 rz -78.89 deg; joints [58.117, 47.637, -22.001, -42.365, -88.704, 135.676]
  MoveL 118 to (283.06, 180.64, 212.36) mm, rotated rx 164.21 ry -43.9 rz -78.89 deg; joints [58.002, 47.885, -21.8, -42.321, -88.924, 135.62]
  MoveL 119 to (282.48, 182.88, 212.36) mm, rotated rx 164.21 ry -43.9 rz -78.89 deg; joints [57.885, 48.13, -21.602, -42.277, -89.144, 135.566]
  MoveL 120 to (282.43, 186.73, 212.36) mm, rotated rx 164.21 ry -43.9 rz -78.89 deg; joints [57.648, 48.436, -21.353, -42.19, -89.477, 135.562]
  MoveL 121 to (283.73, 190.37, 212.36) mm, rotated rx 164.21 ry -43.9 rz -78.89 deg; joints [57.373, 48.563, -21.249, -42.091, -89.726, 135.683]
  MoveL 122 to (286.01, 193.5, 212.36) mm, rotated rx 164.21 ry -43.9 rz -78.89 deg; joints [57.09, 48.53, -21.276, -41.989, -89.882, 135.896]
  MoveL 123 to (288.61, 195.56, 212.36) mm, rotated rx 164.21 ry -43.9 rz -78.89 deg; joints [56.86, 48.375, -21.403, -41.906, -89.931, 136.14]
  MoveL 124 to (291.78, 196.55, 212.36) mm, rotated rx 164.21 ry -43.9 rz -78.89 deg; joints [56.672, 48.067, -21.653, -41.838, -89.862, 136.438]
  MoveL 125 to (295.11, 197, 212.36) mm, rotated rx 164.21 ry -43.9 rz -78.89 deg; joints [56.51, 47.699, -21.951, -41.778, -89.74, 136.749]
  MoveL 126 to (298.46, 197.27, 212.36) mm, rotated rx 164.21 ry -43.9 rz -78.89 deg; joints [56.357, 47.319, -22.257, -41.723, -89.606, 137.058]
  MoveL 127 to (301.81, 197.4, 212.36) mm, rotated rx 164.21 ry -43.9 rz -78.89 deg; joints [56.211, 46.933, -22.568, -41.669, -89.464, 137.366]
  MoveL 128 to (305.16, 197.45, 212.36) mm, rotated rx 164.21 ry -43.9 rz -78.89 deg; joints [56.07, 46.543, -22.88, -41.618, -89.317, 137.67]
  MoveL 129 to (308.51, 197.42, 212.36) mm, rotated rx 164.21 ry -43.9 rz -78.89 deg; joints [55.932, 46.151, -23.191, -41.568, -89.169, 137.972]
  MoveL 130 to (315.39, 197.24, 212.36) mm, rotated rx 164.21 ry -43.9 rz -78.89 deg; joints [55.653, 45.349, -23.824, -41.467, -88.864, 138.583]
  MoveL 131 to (322.27, 197.02, 212.36) mm, rotated rx 164.21 ry -43.9 rz -78.89 deg; joints [55.372, 44.56, -24.441, -41.366, -88.571, 139.183]
  MoveL 132 to (329.11, 197.41, 212.36) mm, rotated rx 164.21 ry -43.9 rz -78.89 deg; joints [55.051, 43.836, -25.002, -41.248, -88.342, 139.773]
  MoveL 133 to (335.99, 199.03, 212.36) mm, rotated rx 164.21 ry -43.9 rz -78.89 deg; joints [54.646, 43.213, -25.48, -41.093, -88.224, 140.363]
  MoveL 134 to (340.16, 199.91, 212.36) mm, rotated rx 164.21 ry -43.9 rz -78.89 deg; joints [54.405, 42.834, -25.769, -41, -88.149, 140.717]
  MoveL 135 to (343.46, 200.32, 212.36) mm, rotated rx 164.21 ry -43.9 rz -78.89 deg; joints [54.23, 42.516, -26.01, -40.932, -88.069, 140.995]
  MoveL 136 to (346, 200.48, 212.36) mm, rotated rx 164.21 ry -43.9 rz -78.89 deg; joints [54.104, 42.26, -26.204, -40.884, -87.997, 141.207]
  MoveL 137 to (348.2, 200.52, 212.36) mm, rotated rx 164.21 ry -43.9 rz -78.89 deg; joints [54.002, 42.033, -26.375, -40.846, -87.928, 141.388]
  MoveL 138 to (350.49, 200.52, 212.36) mm, rotated rx 164.21 ry -43.9 rz -78.89 deg; joints [53.897, 41.794, -26.554, -40.806, -87.854, 141.576]
  MoveL 139 to (352.7, 200.52, 212.36) mm, rotated rx 164.21 ry -43.9 rz -78.89 deg; joints [53.795, 41.564, -26.726, -40.767, -87.783, 141.758]
  MoveL 140 to (355.57, 200.52, 212.36) mm, rotated rx 164.21 ry -43.9 rz -78.89 deg; joints [53.662, 41.269, -26.946, -40.716, -87.693, 141.992]
  MoveL 141 to (359, 200.52, 212.36) mm, rotated rx 164.21 ry -43.9 rz -78.89 deg; joints [53.502, 40.917, -27.206, -40.655, -87.589, 142.27]
  MoveL 142 to (362.6, 200.52, 212.36) mm, rotated rx 164.21 ry -43.9 rz -78.89 deg; joints [53.333, 40.551, -27.477, -40.589, -87.482, 142.56]
  Establecer velocidad (1000.0 mm/s)
  MoveL 143 to (362.6, 200.52, 212.36) mm, rotated rx 164.21 ry -43.9 rz -78.89 deg; joints [53.333, 40.551, -27.477, -40.589, -87.482, 142.56]
  MoveL 144 to (382.21, 200.52, 310.42) mm, rotated rx 164.21 ry -43.9 rz -78.89 deg; joints [52.387, 34.35, -17.597, -40.379, -95.57, 136.815]

--- program pladergr (robot Fanuc LR Mate 200iD/7L) ---
  Suave(1)
  Establecer velocidad (1000.0 mm/s)
  Est. Ref.: RobotiQ 2F-140 Gripper (Mechanism) Base
  Est. herr: Tool 1
  Mostrar Tool 1
  MoveJ 1 to (323.99, 159.18, 238.35) mm, rotated rx 168.3 ry -14.7 rz -86.98 deg; joints [75.345, 48.786, -5.279, -17.745, -78.205, 108.808]
  MoveL 2 to (323.99, 159.18, 238.35) mm, rotated rx 168.3 ry -14.7 rz -86.98 deg; joints [75.345, 48.786, -5.279, -17.745, -78.205, 108.808]
  MoveL 3 to (304.38, 159.18, 140.29) mm, rotated rx 168.3 ry -14.7 rz -86.98 deg; joints [75.692, 53.99, -14.411, -18.538, -69.419, 111.428]
  MoveL 4 to (304.38, 159.18, 140.29) mm, rotated rx 168.3 ry -14.7 rz -86.98 deg; joints [75.692, 53.99, -14.411, -18.538, -69.419, 111.428]
  Establecer velocidad (50.0 mm/s)
  MoveL 5 to (318.28, 160.81, 140.29) mm, rotated rx 168.3 ry -14.7 rz -86.98 deg; joints [75.336, 51.733, -16.323, -18.811, -67.717, 112.434]
  MoveL 6 to (332.27, 160.99, 140.29) mm, rotated rx 168.3 ry -14.7 rz -86.98 deg; joints [75.069, 49.552, -18.125, -19.085, -66.095, 113.333]
  MoveL 7 to (346.25, 160.87, 140.29) mm, rotated rx 168.3 ry -14.7 rz -86.98 deg; joints [74.813, 47.483, -19.795, -19.359, -64.599, 114.189]
  MoveL 8 to (360.2, 160.1, 140.52) mm, rotated rx 168.3 ry -14.7 rz -86.98 deg; joints [74.596, 45.483, -21.335, -19.628, -63.215, 114.975]
  MoveL 9 to (374.69, 158.54, 142.06) mm, rotated rx 168.3 ry -14.7 rz -86.98 deg; joints [74.418, 43.406, -22.706, -19.882, -61.98, 115.672]
  MoveL 10 to (388.82, 156.24, 144.98) mm, rotated rx 168.3 ry -14.7 rz -86.98 deg; joints [74.296, 41.353, -23.811, -20.096, -60.98, 116.222]
  MoveL 11 to (402.6, 153.26, 149.26) mm, rotated rx 168.3 ry -14.7 rz -86.98 deg; joints [74.228, 39.305, -24.661, -20.266, -60.204, 116.625]
  MoveL 12 to (416.24, 149.6, 153.81) mm, rotated rx 168.3 ry -14.7 rz -86.98 deg; joints [74.214, 37.275, -25.401, -20.417, -59.514, 116.937]
  MoveL 13 to (430.22, 146.2, 157.02) mm, rotated rx 168.3 ry -14.7 rz -86.98 deg; joints [74.17, 35.309, -26.236, -20.595, -58.746, 117.32]
  MoveL 14 to (444.55, 143.57, 158.87) mm, rotated rx 168.3 ry -14.7 rz -86.98 deg; joints [74.054, 33.422, -27.163, -20.804, -57.916, 117.819]
  MoveL 15 to (460.25, 141.64, 159.34) mm, rotated rx 168.3 ry -14.7 rz -86.98 deg; joints [73.843, 31.498, -28.265, -21.069, -56.953, 118.493]
  MoveL 16 to (476.08, 140.69, 159.34) mm, rotated rx 168.3 ry -14.7 rz -86.98 deg; joints [73.536, 29.648, -29.34, -21.345, -56.047, 119.261]
  MoveL 17 to (491.93, 140.58, 159.34) mm, rotated rx 168.3 ry -14.7 rz -86.98 deg; joints [73.141, 27.849, -30.338, -21.616, -55.245, 120.089]
  MoveL 18 to (507.79, 140.58, 159.34) mm, rotated rx 168.3 ry -14.7 rz -86.98 deg; joints [72.716, 26.075, -31.272, -21.88, -54.512, 120.927]
  MoveL 19 to (523.64, 140.58, 159.34) mm, rotated rx 168.3 ry -14.7 rz -86.98 deg; joints [72.271, 24.319, -32.147, -22.136, -53.843, 121.765]
  MoveL 20 to (563.28, 140.58, 159.34) mm, rotated rx 168.3 ry -14.7 rz -86.98 deg; joints [71.054, 19.981, -34.087, -22.733, -52.438, 123.868]
  MoveL 21 to (570.04, 140.04, 159.34) mm, rotated rx 168.3 ry -14.7 rz -86.98 deg; joints [70.881, 19.225, -34.391, -22.828, -52.214, 124.182]
  MoveL 22 to (576.96, 137.96, 159.34) mm, rotated rx 168.3 ry -14.7 rz -86.98 deg; joints [70.85, 18.394, -34.714, -22.927, -51.926, 124.371]
  MoveL 23 to (583.51, 134.22, 159.34) mm, rotated rx 168.3 ry -14.7 rz -86.98 deg; joints [70.995, 17.539, -35.032, -23.021, -51.587, 124.39]
  MoveL 24 to (589.11, 128.98, 159.34) mm, rotated rx 168.3 ry -14.7 rz -86.98 deg; joints [71.328, 16.732, -35.319, -23.103, -51.216, 124.214]
  MoveL 25 to (593.3, 122.66, 159.34) mm, rotated rx 168.3 ry -14.7 rz -86.98 deg; joints [71.827, 16.042, -35.556, -23.165, -50.839, 123.852]
  MoveL 26 to (595.85, 115.8, 159.34) mm, rotated rx 168.3 ry -14.7 rz -86.98 deg; joints [72.446, 15.518, -35.729, -23.203, -50.481, 123.342]
  MoveL 27 to (596.8, 108.99, 159.34) mm, rotated rx 168.3 ry -14.7 rz -86.98 deg; joints [73.123, 15.18, -35.838, -23.215, -50.165, 122.743]
  MoveL 28 to (596.82, 102.38, 159.34) mm, rotated rx 168.3 ry -14.7 rz -86.98 deg; joints [73.813, 14.96, -35.908, -23.212, -49.88, 122.108]
  MoveL 29 to (596.79, 95.78, 159.34) mm, rotated rx 168.3 ry -14.7 rz -86.98 deg; joints [74.51, 14.753, -35.972, -23.203, -49.599, 121.462]
  MoveL 30 to (595.8, 88.96, 159.34) mm, rotated rx 168.3 ry -14.7 rz -86.98 deg; joints [75.261, 14.658, -36.002, -23.177, -49.332, 120.742]
  MoveL 31 to (593.21, 82.11, 159.34) mm, rotated rx 168.3 ry -14.7 rz -86.98 deg; joints [76.059, 14.753, -35.972, -23.124, -49.105, 119.942]
  MoveL 32 to (588.98, 75.81, 159.34) mm, rotated rx 168.3 ry -14.7 rz -86.98 deg; joints [76.838, 15.059, -35.876, -23.044, -48.947, 119.124]
  MoveL 33 to (583.34, 70.6, 159.34) mm, rotated rx 168.3 ry -14.7 rz -86.98 deg; joints [77.525, 15.562, -35.714, -22.943, -48.878, 118.36]
  MoveL 34 to (576.77, 66.91, 159.34) mm, rotated rx 168.3 ry -14.7 rz -86.98 deg; joints [78.063, 16.215, -35.497, -22.831, -48.908, 117.712]
  MoveL 35 to (568.86, 64.71, 159.34) mm, rotated rx 168.3 ry -14.7 rz -86.98 deg; joints [78.462, 17.058, -35.204, -22.702, -49.052, 117.164]
  MoveL 36 to (561.21, 64.37, 159.34) mm, rotated rx 168.3 ry -14.7 rz -86.98 deg; joints [78.657, 17.915, -34.893, -22.584, -49.278, 116.812]
  MoveL 37 to (553.66, 64.37, 159.34) mm, rotated rx 168.3 ry -14.7 rz -86.98 deg; joints [78.809, 18.768, -34.569, -22.465, -49.529, 116.496]
  MoveL 38 to (546.11, 64.37, 159.34) mm, rotated rx 168.3 ry -14.7 rz -86.98 deg; joints [78.958, 19.62, -34.233, -22.344, -49.793, 116.179]
  MoveL 39 to (538.56, 64.37, 159.34) mm, rotated rx 168.3 ry -14.7 rz -86.98 deg; joints [79.102, 20.473, -33.883, -22.22, -50.072, 115.861]
  MoveL 40 to (531.01, 64.37, 159.34) mm, rotated rx 168.3 ry -14.7 rz -86.98 deg; joints [79.243, 21.327, -33.52, -22.094, -50.364, 115.541]
  MoveL 41 to (523.46, 64.37, 159.34) mm, rotated rx 168.3 ry -14.7 rz -86.98 deg; joints [79.381, 22.181, -33.143, -21.965, -50.67, 115.22]
  MoveL 42 to (506.02, 64.37, 159.34) mm, rotated rx 168.3 ry -14.7 rz -86.98 deg; joints [79.685, 24.161, -32.223, -21.661, -51.429, 114.474]
  MoveL 43 to (488.58, 64.37, 159.34) mm, rotated rx 168.3 ry -14.7 rz -86.98 deg; joints [79.973, 26.155, -31.23, -21.347, -52.263, 113.722]
  MoveL 44 to (471.15, 64.63, 159.34) mm, rotated rx 168.3 ry -14.7 rz -86.98 deg; joints [80.223, 28.172, -30.161, -21.028, -53.182, 112.985]
  MoveL 45 to (453.71, 64.24, 159.32) mm, rotated rx 168.3 ry -14.7 rz -86.98 deg; joints [80.514, 30.203, -29.025, -20.7, -54.153, 112.189]
  MoveL 46 to (439.06, 63.09, 158.33) mm, rotated rx 168.3 ry -14.7 rz -86.98 deg; joints [80.818, 31.97, -28.131, -20.444, -54.897, 111.497]
  MoveL 47 to (424.75, 61.24, 155.94) mm, rotated rx 168.3 ry -14.7 rz -86.98 deg; joints [81.162, 33.778, -27.371, -20.222, -55.503, 110.827]
  MoveL 48 to (410.78, 58.72, 152.16) mm, rotated rx 168.3 ry -14.7 rz -86.98 deg; joints [81.543, 35.626, -26.739, -20.03, -55.98, 110.179]
  MoveL 49 to (397.11, 55.55, 147.38) mm, rotated rx 168.3 ry -14.7 rz -86.98 deg; joints [81.958, 37.502, -26.183, -19.854, -56.376, 109.53]
  MoveL 50 to (383.35, 51.64, 143.68) mm, rotated rx 168.3 ry -14.7 rz -86.98 deg; joints [82.417, 39.351, -25.437, -19.632, -56.939, 108.762]
  MoveL 51 to (369.48, 46.98, 141.34) mm, rotated rx 168.3 ry -14.7 rz -86.98 deg; joints [82.918, 41.176, -24.464, -19.361, -57.705, 107.868]
  MoveL 52 to (354.24, 42.7, 140.31) mm, rotated rx 168.3 ry -14.7 rz -86.98 deg; joints [83.385, 43.181, -23.125, -19.027, -58.828, 106.876]
  MoveL 53 to (338.6, 39.9, 140.29) mm, rotated rx 168.3 ry -14.7 rz -86.98 deg; joints [83.728, 45.299, -21.51, -18.674, -60.254, 105.922]
  MoveL 54 to (322.7, 38.61, 140.29) mm, rotated rx 168.3 ry -14.7 rz -86.98 deg; joints [83.95, 47.579, -19.717, -18.329, -61.889, 105.048]
  MoveL 55 to (306.75, 38.86, 140.29) mm, rotated rx 168.3 ry -14.7 rz -86.98 deg; joints [84.052, 50.025, -17.737, -17.997, -63.74, 104.25]
  MoveL 56 to (290.97, 40.63, 140.37) mm, rotated rx 168.3 ry -14.7 rz -86.98 deg; joints [84.043, 52.643, -15.546, -17.683, -65.829, 103.518]
  MoveL 57 to (281.29, 42.5, 140.79) mm, rotated rx 168.3 ry -14.7 rz -86.98 deg; joints [83.983, 54.366, -14.02, -17.491, -67.301, 103.075]
  MoveL 58 to (271.77, 44.93, 141.55) mm, rotated rx 168.3 ry -14.7 rz -86.98 deg; joints [83.886, 56.176, -12.345, -17.304, -68.927, 102.633]
  MoveL 59 to (262.4, 47.92, 142.63) mm, rotated rx 168.3 ry -14.7 rz -86.98 deg; joints [83.751, 58.109, -10.489, -17.122, -70.739, 102.182]
  MoveL 60 to (253.55, 52.02, 143.98) mm, rotated rx 168.3 ry -14.7 rz -86.98 deg; joints [83.542, 60.149, -8.472, -16.958, -72.728, 101.768]
  MoveL 61 to (245.67, 57.8, 145.44) mm, rotated rx 168.3 ry -14.7 rz -86.98 deg; joints [83.218, 62.249, -6.35, -16.826, -74.851, 101.445]
  MoveL 62 to (239.11, 64.99, 146.84) mm, rotated rx 168.3 ry -14.7 rz -86.98 deg; joints [82.798, 64.347, -4.203, -16.732, -77.028, 101.219]
  MoveL 63 to (234.07, 73.41, 148.04) mm, rotated rx 168.3 ry -14.7 rz -86.98 deg; joints [82.292, 66.385, -2.105, -16.68, -79.183, 101.097]
  MoveL 64 to (230.81, 82.64, 148.87) mm, rotated rx 168.3 ry -14.7 rz -86.98 deg; joints [81.724, 68.198, -0.242, -16.67, -81.13, 101.107]
  MoveL 65 to (229.67, 89.16, 149.17) mm, rotated rx 168.3 ry -14.7 rz -86.98 deg; joints [81.315, 69.173, 0.751, -16.687, -82.199, 101.215]
  MoveL 66 to (229.4, 95.77, 149.25) mm, rotated rx 168.3 ry -14.7 rz -86.98 deg; joints [80.893, 69.837, 1.413, -16.723, -82.955, 101.431]
  MoveL 67 to (229.51, 102.4, 149.22) mm, rotated rx 168.3 ry -14.7 rz -86.98 deg; joints [80.467, 70.37, 1.936, -16.766, -83.578, 101.689]
  MoveL 68 to (230.74, 108.84, 148.89) mm, rotated rx 168.3 ry -14.7 rz -86.98 deg; joints [80.042, 70.279, 1.802, -16.83, -83.572, 102.138]
  MoveL 69 to (234.4, 116.78, 147.96) mm, rotated rx 168.3 ry -14.7 rz -86.98 deg; joints [79.492, 69.087, 0.501, -16.951, -82.487, 103.049]
  MoveL 70 to (239.88, 123.56, 146.67) mm, rotated rx 168.3 ry -14.7 rz -86.98 deg; joints [78.991, 67.269, -1.442, -17.101, -80.776, 104.108]
  MoveL 71 to (245.96, 129.74, 145.38) mm, rotated rx 168.3 ry -14.7 rz -86.98 deg; joints [78.516, 65.537, -3.276, -17.258, -79.164, 105.118]
  MoveL 72 to (255.89, 138.09, 143.59) mm, rotated rx 168.3 ry -14.7 rz -86.98 deg; joints [77.842, 63.108, -5.805, -17.5, -76.952, 106.546]
  MoveL 73 to (266.81, 145.34, 142.08) mm, rotated rx 168.3 ry -14.7 rz -86.98 deg; joints [77.213, 60.774, -8.162, -17.752, -74.893, 107.895]
  MoveL 74 to (278.5, 151.29, 140.97) mm, rotated rx 168.3 ry -14.7 rz -86.98 deg; joints [76.644, 58.513, -10.357, -18.008, -72.977, 109.153]
  MoveL 75 to (290.78, 155.88, 140.37) mm, rotated rx 168.3 ry -14.7 rz -86.98 deg; joints [76.142, 56.304, -12.395, -18.265, -71.193, 110.31]
  Establecer velocidad (1000.0 mm/s)
  MoveL 76 to (290.78, 155.88, 140.37) mm, rotated rx 168.3 ry -14.7 rz -86.98 deg; joints [76.142, 56.304, -12.395, -18.265, -71.193, 110.31]
  MoveL 77 to (310.4, 155.88, 238.43) mm, rotated rx 168.3 ry -14.7 rz -86.98 deg; joints [75.812, 51.316, -3.243, -17.576, -80.004, 107.727]
  Establecer velocidad (1000.0 mm/s)
  MoveL 78 to (543.44, 140.78, 316.08) mm, rotated rx 168.3 ry -14.7 rz -86.98 deg; joints [71.663, 15.752, -12.896, -18.713, -72.105, 114.845]
  MoveL 79 to (523.83, 140.78, 218.03) mm, rotated rx 168.3 ry -14.7 rz -86.98 deg; joints [72.247, 21.232, -24.792, -20.42, -60.707, 118.617]
  MoveL 80 to (523.83, 140.78, 218.03) mm, rotated rx 168.3 ry -14.7 rz -86.98 deg; joints [72.247, 21.232, -24.792, -20.42, -60.707, 118.617]
  Establecer velocidad (50.0 mm/s)
  MoveL 81 to (547.65, 139.64, 218.03) mm, rotated rx 168.3 ry -14.7 rz -86.98 deg; joints [71.639, 18.427, -25.852, -20.665, -59.906, 119.637]
  MoveL 82 to (571.28, 136.35, 218.03) mm, rotated rx 168.3 ry -14.7 rz -86.98 deg; joints [71.197, 15.578, -26.787, -20.882, -59.172, 120.452]
  MoveL 83 to (578.97, 134.27, 218.03) mm, rotated rx 168.3 ry -14.7 rz -86.98 deg; joints [71.144, 14.612, -27.071, -20.946, -58.924, 120.621]
  MoveL 84 to (585.97, 130.56, 218.03) mm, rotated rx 168.3 ry -14.7 rz -86.98 deg; joints [71.276, 13.66, -27.333, -20.996, -58.637, 120.603]
  MoveL 85 to (592.06, 125.43, 218.03) mm, rotated rx 168.3 ry -14.7 rz -86.98 deg; joints [71.586, 12.759, -27.566, -21.033, -58.321, 120.399]
  MoveL 86 to (596.85, 119.1, 218.03) mm, rotated rx 168.3 ry -14.7 rz -86.98 deg; joints [72.073, 11.962, -27.76, -21.052, -57.986, 120.007]
  MoveL 87 to (599.88, 111.76, 218.03) mm, rotated rx 168.3 ry -14.7 rz -86.98 deg; joints [72.735, 11.338, -27.902, -21.05, -57.643, 119.423]
  MoveL 88 to (600.77, 103.88, 218.03) mm, rotated rx 168.3 ry -14.7 rz -86.98 deg; joints [73.534, 10.955, -27.987, -21.023, -57.31, 118.677]
  MoveL 89 to (600.39, 95.98, 218.03) mm, rotated rx 168.3 ry -14.7 rz -86.98 deg; joints [74.382, 10.732, -28.034, -20.981, -56.998, 117.866]
  MoveL 90 to (598.12, 88.46, 218.03) mm, rotated rx 168.3 ry -14.7 rz -86.98 deg; joints [75.249, 10.758, -28.028, -20.921, -56.73, 117.01]
  MoveL 91 to (593.96, 81.74, 218.03) mm, rotated rx 168.3 ry -14.7 rz -86.98 deg; joints [76.078, 11.049, -27.966, -20.845, -56.527, 116.164]
  MoveL 92 to (588.43, 76.11, 218.03) mm, rotated rx 168.3 ry -14.7 rz -86.98 deg; joints [76.818, 11.546, -27.855, -20.76, -56.398, 115.383]
  MoveL 93 to (582.02, 71.88, 218.03) mm, rotated rx 168.3 ry -14.7 rz -86.98 deg; joints [77.42, 12.194, -27.704, -20.674, -56.351, 114.721]
  MoveL 94 to (574.85, 69.17, 218.03) mm, rotated rx 168.3 ry -14.7 rz -86.98 deg; joints [77.869, 12.977, -27.511, -20.589, -56.392, 114.192]
  MoveL 95 to (567.36, 67.81, 218.03) mm, rotated rx 168.3 ry -14.7 rz -86.98 deg; joints [78.175, 13.835, -27.286, -20.509, -56.507, 113.792]
  MoveL 96 to (559.81, 66.71, 218.03) mm, rotated rx 168.3 ry -14.7 rz -86.98 deg; joints [78.447, 14.707, -27.043, -20.427, -56.65, 113.419]
  MoveL 97 to (540.48, 64.87, 218.03) mm, rotated rx 168.3 ry -14.7 rz -86.98 deg; joints [79.017, 16.967, -26.349, -20.215, -57.124, 112.561]
  MoveL 98 to (521.07, 64.35, 218.03) mm, rotated rx 168.3 ry -14.7 rz -86.98 deg; joints [79.426, 19.274, -25.546, -19.997, -57.752, 111.824]
  MoveL 99 to (503.42, 64.87, 218.03) mm, rotated rx 168.3 ry -14.7 rz -86.98 deg; joints [79.682, 21.404, -24.721, -19.795, -58.448, 111.236]
  MoveL 100 to (485.95, 66.81, 218.03) mm, rotated rx 168.3 ry -14.7 rz -86.98 deg; joints [79.794, 23.56, -23.809, -19.597, -59.273, 110.764]
  MoveL 101 to (468.82, 70.05, 218.03) mm, rotated rx 168.3 ry -14.7 rz -86.98 deg; joints [79.78, 25.724, -22.815, -19.405, -60.214, 110.394]
  MoveL 102 to (451.38, 69.87, 218.03) mm, rotated rx 168.3 ry -14.7 rz -86.98 deg; joints [80.065, 27.881, -21.75, -19.176, -61.132, 109.705]
  MoveL 103 to (433.94, 69.77, 218.03) mm, rotated rx 168.3 ry -14.7 rz -86.98 deg; joints [80.328, 30.079, -20.591, -18.941, -62.147, 109.012]
  MoveL 104 to (428.75, 69.89, 218.03) mm, rotated rx 168.3 ry -14.7 rz -86.98 deg; joints [80.391, 30.745, -20.226, -18.872, -62.474, 108.815]
  MoveL 105 to (423.57, 70.15, 218.03) mm, rotated rx 168.3 ry -14.7 rz -86.98 deg; joints [80.442, 31.417, -19.85, -18.803, -62.814, 108.628]
  MoveL 106 to (418.4, 70.59, 218.03) mm, rotated rx 168.3 ry -14.7 rz -86.98 deg; joints [80.477, 32.097, -19.464, -18.736, -63.169, 108.453]
  MoveL 107 to (413.29, 71.43, 218.03) mm, rotated rx 168.3 ry -14.7 rz -86.98 deg; joints [80.478, 32.783, -19.067, -18.672, -63.545, 108.31]
  MoveL 108 to (408.77, 73.9, 218.03) mm, rotated rx 168.3 ry -14.7 rz -86.98 deg; joints [80.34, 33.434, -18.684, -18.628, -63.949, 108.311]
  MoveL 109 to (405.82, 77.05, 218.03) mm, rotated rx 168.3 ry -14.7 rz -86.98 deg; joints [80.128, 33.897, -18.408, -18.61, -64.275, 108.425]
  MoveL 110 to (403.89, 80.91, 218.03) mm, rotated rx 168.3 ry -14.7 rz -86.98 deg; joints [79.847, 34.244, -18.199, -18.611, -64.558, 108.631]
  MoveL 111 to (403.34, 85.17, 218.03) mm, rotated rx 168.3 ry -14.7 rz -86.98 deg; joints [79.515, 34.422, -18.092, -18.633, -64.76, 108.924]
  MoveL 112 to (404.24, 89.4, 218.03) mm, rotated rx 168.3 ry -14.7 rz -86.98 deg; joints [79.166, 34.407, -18.101, -18.674, -64.858, 109.275]
  MoveL 113 to (405.62, 93.52, 218.03) mm, rotated rx 168.3 ry -14.7 rz -86.98 deg; joints [78.817, 34.33, -18.148, -18.719, -64.92, 109.638]
  MoveL 114 to (407.03, 97.64, 218.03) mm, rotated rx 168.3 ry -14.7 rz -86.98 deg; joints [78.469, 34.252, -18.195, -18.764, -64.982, 110.001]
  MoveL 115 to (407.43, 100.93, 218.03) mm, rotated rx 168.3 ry -14.7 rz -86.98 deg; joints [78.201, 34.29, -18.172, -18.789, -65.085, 110.259]
  MoveL 116 to (406.44, 104.27, 218.03) mm, rotated rx 168.3 ry -14.7 rz -86.98 deg; joints [77.954, 34.515, -18.036, -18.795, -65.29, 110.455]
  MoveL 117 to (405.47, 107.61, 218.03) mm, rotated rx 168.3 ry -14.7 rz -86.98 deg; joints [77.707, 34.74, -17.899, -18.801, -65.495, 110.651]
  MoveL 118 to (404.52, 110.96, 218.03) mm, rotated rx 168.3 ry -14.7 rz -86.98 deg; joints [77.46, 34.964, -17.761, -18.806, -65.701, 110.847]
  MoveL 119 to (403.64, 114.32, 218.03) mm, rotated rx 168.3 ry -14.7 rz -86.98 deg; joints [77.212, 35.183, -17.627, -18.811, -65.905, 111.044]
  MoveL 120 to (403.58, 120.1, 218.03) mm, rotated rx 168.3 ry -14.7 rz -86.98 deg; joints [76.762, 35.37, -17.511, -18.84, -66.153, 111.448]
  MoveL 121 to (405.52, 125.56, 218.03) mm, rotated rx 168.3 ry -14.7 rz -86.98 deg; joints [76.3, 35.285, -17.564, -18.892, -66.245, 111.922]
  MoveL 122 to (408.94, 130.25, 218.03) mm, rotated rx 168.3 ry -14.7 rz -86.98 deg; joints [75.869, 34.984, -17.749, -18.959, -66.203, 112.412]
  MoveL 123 to (412.84, 133.34, 218.03) mm, rotated rx 168.3 ry -14.7 rz -86.98 deg; joints [75.551, 34.573, -18, -19.024, -66.064, 112.815]
  MoveL 124 to (417.59, 134.83, 218.03) mm, rotated rx 168.3 ry -14.7 rz -86.98 deg; joints [75.337, 34, -18.347, -19.093, -65.803, 113.149]
  MoveL 125 to (422.59, 135.5, 218.03) mm, rotated rx 168.3 ry -14.7 rz -86.98 deg; joints [75.181, 33.373, -18.721, -19.163, -65.498, 113.437]
  MoveL 126 to (427.61, 135.9, 218.03) mm, rotated rx 168.3 ry -14.7 rz -86.98 deg; joints [75.043, 32.738, -19.094, -19.231, -65.189, 113.707]
  MoveL 127 to (432.64, 136.11, 218.03) mm, rotated rx 168.3 ry -14.7 rz -86.98 deg; joints [74.919, 32.102, -19.461, -19.298, -64.88, 113.963]
  MoveL 128 to (437.66, 136.17, 218.03) mm, rotated rx 168.3 ry -14.7 rz -86.98 deg; joints [74.805, 31.466, -19.823, -19.364, -64.574, 114.207]
  MoveL 129 to (442.69, 136.13, 218.03) mm, rotated rx 168.3 ry -14.7 rz -86.98 deg; joints [74.698, 30.831, -20.179, -19.429, -64.273, 114.444]
  MoveL 130 to (453.01, 135.86, 218.03) mm, rotated rx 168.3 ry -14.7 rz -86.98 deg; joints [74.488, 29.534, -20.886, -19.561, -63.672, 114.913]
  MoveL 131 to (463.33, 135.53, 218.03) mm, rotated rx 168.3 ry -14.7 rz -86.98 deg; joints [74.277, 28.252, -21.561, -19.691, -63.102, 115.374]
  MoveL 132 to (473.59, 136.11, 218.03) mm, rotated rx 168.3 ry -14.7 rz -86.98 deg; joints [73.983, 27.023, -22.183, -19.821, -62.608, 115.898]
  MoveL 133 to (483.91, 138.54, 218.03) mm, rotated rx 168.3 ry -14.7 rz -86.98 deg; joints [73.522, 25.865, -22.748, -19.955, -62.222, 116.568]
  MoveL 134 to (490.17, 139.86, 218.03) mm, rotated rx 168.3 ry -14.7 rz -86.98 deg; joints [73.248, 25.164, -23.08, -20.034, -61.996, 116.964]
  MoveL 135 to (495.12, 140.48, 218.03) mm, rotated rx 168.3 ry -14.7 rz -86.98 deg; joints [73.065, 24.597, -23.342, -20.094, -61.808, 117.245]
  MoveL 136 to (498.93, 140.72, 218.03) mm, rotated rx 168.3 ry -14.7 rz -86.98 deg; joints [72.943, 24.153, -23.544, -20.139, -61.657, 117.443]
  MoveL 137 to (502.22, 140.78, 218.03) mm, rotated rx 168.3 ry -14.7 rz -86.98 deg; joints [72.85, 23.766, -23.718, -20.177, -61.523, 117.602]
  MoveL 138 to (505.66, 140.78, 218.03) mm, rotated rx 168.3 ry -14.7 rz -86.98 deg; joints [72.757, 23.361, -23.896, -20.217, -61.385, 117.764]
  MoveL 139 to (508.99, 140.78, 218.03) mm, rotated rx 168.3 ry -14.7 rz -86.98 deg; joints [72.665, 22.97, -24.067, -20.255, -61.254, 117.92]
  MoveL 140 to (513.28, 140.78, 218.03) mm, rotated rx 168.3 ry -14.7 rz -86.98 deg; joints [72.546, 22.465, -24.282, -20.303, -61.089, 118.122]
  MoveL 141 to (518.42, 140.78, 218.03) mm, rotated rx 168.3 ry -14.7 rz -86.98 deg; joints [72.402, 21.863, -24.534, -20.361, -60.899, 118.363]
  MoveL 142 to (523.83, 140.78, 218.03) mm, rotated rx 168.3 ry -14.7 rz -86.98 deg; joints [72.247, 21.232, -24.792, -20.42, -60.707, 118.617]
  Establecer velocidad (1000.0 mm/s)
  MoveL 143 to (523.83, 140.78, 218.03) mm, rotated rx 168.3 ry -14.7 rz -86.98 deg; joints [72.247, 21.232, -24.792, -20.42, -60.707, 118.617]
  MoveL 144 to (543.44, 140.78, 316.08) mm, rotated rx 168.3 ry -14.7 rz -86.98 deg; joints [71.663, 15.752, -12.896, -18.713, -72.105, 114.845]

--- program arrizch (robot Fanuc LR Mate 200iD/7L) ---
  Suave(1)
  Establecer velocidad (1000.0 mm/s)
  Est. Ref.: RobotiQ 2F-140 Gripper (Mechanism) Base
  Est. herr: Tool 1
  Mostrar Tool 1
  MoveJ 1 to (227.79, -210.8, 228.5) mm, rotated rx 167 ry 29.36 rz -96.45 deg; joints [112.467, 45.334, -15.632, 32.503, -78.699, 56.721]
  MoveL 2 to (227.79, -210.8, 228.5) mm, rotated rx 167 ry 29.36 rz -96.45 deg; joints [112.467, 45.334, -15.632, 32.503, -78.699, 56.721]
  MoveL 3 to (208.18, -210.8, 130.44) mm, rotated rx 167 ry 29.36 rz -96.45 deg; joints [111.928, 52.063, -23.982, 33.793, -71.427, 52.439]
  MoveL 4 to (208.18, -210.8, 130.44) mm, rotated rx 167 ry 29.36 rz -96.45 deg; joints [111.928, 52.063, -23.982, 33.793, -71.427, 52.439]
  Establecer velocidad (50.0 mm/s)
  MoveL 5 to (200.4, -210.8, 129.52) mm, rotated rx 167 ry 29.36 rz -96.45 deg; joints [111.72, 53.181, -23.134, 33.668, -72.026, 53.101]
  MoveL 6 to (192.62, -210.8, 128.43) mm, rotated rx 167 ry 29.36 rz -96.45 deg; joints [111.516, 54.34, -22.264, 33.544, -72.646, 53.771]
  MoveL 7 to (184.01, -210.8, 127.03) mm, rotated rx 167 ry 29.36 rz -96.45 deg; joints [111.295, 55.674, -21.269, 33.406, -73.363, 54.524]
  MoveL 8 to (174.28, -210.8, 125.2) mm, rotated rx 167 ry 29.36 rz -96.45 deg; joints [111.05, 57.255, -20.098, 33.249, -74.216, 55.394]
  MoveL 9 to (165.95, -210.8, 123.42) mm, rotated rx 167 ry 29.36 rz -96.45 deg; joints [110.844, 58.679, -19.045, 33.115, -74.991, 56.16]
  MoveL 10 to (162, -210.8, 122.51) mm, rotated rx 167 ry 29.36 rz -96.45 deg; joints [110.748, 59.378, -18.527, 33.051, -75.375, 56.531]
  MoveL 11 to (158.5, -210.8, 121.66) mm, rotated rx 167 ry 29.36 rz -96.45 deg; joints [110.664, 60.015, -18.056, 32.994, -75.726, 56.865]
  MoveL 12 to (157.03, -210.8, 121.23) mm, rotated rx 167 ry 29.36 rz -96.45 deg; joints [110.628, 60.289, -17.86, 32.971, -75.872, 57.004]
  MoveL 13 to (156.08, -210.8, 120.61) mm, rotated rx 167 ry 29.36 rz -96.45 deg; joints [110.606, 60.482, -17.767, 32.96, -75.939, 57.075]
  MoveL 14 to (155.28, -210.8, 119.56) mm, rotated rx 167 ry 29.36 rz -96.45 deg; joints [110.586, 60.669, -17.739, 32.958, -75.952, 57.107]
  MoveL 15 to (154.93, -210.8, 118.56) mm, rotated rx 167 ry 29.36 rz -96.45 deg; joints [110.578, 60.774, -17.781, 32.965, -75.912, 57.09]
  MoveL 16 to (154.87, -210.8, 117.34) mm, rotated rx 167 ry 29.36 rz -96.45 deg; joints [110.577, 60.838, -17.892, 32.98, -75.819, 57.029]
  MoveL 17 to (154.87, -210.8, 115.68) mm, rotated rx 167 ry 29.36 rz -96.45 deg; joints [110.577, 60.911, -18.055, 33.003, -75.683, 56.938]
  MoveL 18 to (154.87, -210.8, 112.74) mm, rotated rx 167 ry 29.36 rz -96.45 deg; joints [110.577, 61.043, -18.342, 33.043, -75.442, 56.776]
  MoveL 19 to (154.87, -210.8, 109.33) mm, rotated rx 167 ry 29.36 rz -96.45 deg; joints [110.577, 61.198, -18.672, 33.09, -75.165, 56.59]
  MoveL 20 to (154.87, -210.8, 105.92) mm, rotated rx 167 ry 29.36 rz -96.45 deg; joints [110.577, 61.358, -19, 33.138, -74.89, 56.404]
  MoveL 21 to (154.87, -210.8, 102.42) mm, rotated rx 167 ry 29.36 rz -96.45 deg; joints [110.577, 61.524, -19.334, 33.188, -74.61, 56.215]
  Establecer velocidad (1000.0 mm/s)
  MoveL 22 to (154.87, -210.8, 102.42) mm, rotated rx 167 ry 29.36 rz -96.45 deg; joints [110.577, 61.524, -19.334, 33.188, -74.61, 56.215]
  MoveL 23 to (174.49, -210.8, 200.47) mm, rotated rx 167 ry 29.36 rz -96.45 deg; joints [111.054, 54.52, -12.066, 32.291, -80.975, 59.839]
  Establecer velocidad (1000.0 mm/s)
  MoveL 24 to (235.63, -210.8, 229.26) mm, rotated rx 167 ry 29.36 rz -96.45 deg; joints [112.691, 44.202, -16.375, 32.56, -78.188, 56.128]
  MoveL 25 to (216.02, -210.8, 131.2) mm, rotated rx 167 ry 29.36 rz -96.45 deg; joints [112.141, 50.974, -24.816, 33.919, -70.841, 51.777]
  MoveL 26 to (216.02, -210.8, 131.2) mm, rotated rx 167 ry 29.36 rz -96.45 deg; joints [112.141, 50.974, -24.816, 33.919, -70.841, 51.777]
  Establecer velocidad (50.0 mm/s)
  MoveL 27 to (230.82, -210.8, 133.22) mm, rotated rx 167 ry 29.36 rz -96.45 deg; joints [112.554, 48.958, -26.247, 34.137, -69.864, 50.599]
  MoveL 28 to (247.08, -210.8, 137.18) mm, rotated rx 167 ry 29.36 rz -96.45 deg; joints [113.025, 46.735, -27.523, 34.323, -69.046, 49.462]
  MoveL 29 to (262.81, -210.8, 142.89) mm, rotated rx 167 ry 29.36 rz -96.45 deg; joints [113.498, 44.547, -28.455, 34.439, -68.512, 48.527]
  MoveL 30 to (277.82, -210.8, 150.28) mm, rotated rx 167 ry 29.36 rz -96.45 deg; joints [113.968, 42.397, -29.045, 34.48, -68.259, 47.803]
  MoveL 31 to (291.94, -210.8, 159.28) mm, rotated rx 167 ry 29.36 rz -96.45 deg; joints [114.425, 40.296, -29.294, 34.444, -68.28, 47.297]
  MoveL 32 to (304.98, -210.8, 169.76) mm, rotated rx 167 ry 29.36 rz -96.45 deg; joints [114.863, 38.257, -29.209, 34.336, -68.566, 47.009]
  MoveL 33 to (316.81, -210.8, 181.6) mm, rotated rx 167 ry 29.36 rz -96.45 deg; joints [115.273, 36.302, -28.799, 34.163, -69.107, 46.939]
  Establecer velocidad (1000.0 mm/s)
  MoveL 34 to (316.81, -210.8, 181.6) mm, rotated rx 167 ry 29.36 rz -96.45 deg; joints [115.273, 36.302, -28.799, 34.163, -69.107, 46.939]
  MoveL 35 to (336.42, -210.8, 279.66) mm, rotated rx 167 ry 29.36 rz -96.45 deg; joints [115.98, 29.779, -18.615, 32.383, -77.983, 52.194]
  Establecer velocidad (1000.0 mm/s)
  MoveL 36 to (423.45, -210.8, 252.17) mm, rotated rx 167 ry 29.36 rz -96.45 deg; joints [119.621, 21.243, -26.574, 32.821, -73.086, 44.842]
  MoveL 37 to (403.83, -210.8, 154.11) mm, rotated rx 167 ry 29.36 rz -96.45 deg; joints [118.722, 29.104, -37.674, 35.542, -63.466, 38.815]
  MoveL 38 to (403.83, -210.8, 154.11) mm, rotated rx 167 ry 29.36 rz -96.45 deg; joints [118.722, 29.104, -37.674, 35.542, -63.466, 38.815]
  Establecer velocidad (50.0 mm/s)
  MoveL 39 to (405.69, -210.8, 141.37) mm, rotated rx 167 ry 29.36 rz -96.45 deg; joints [118.805, 29.852, -39.295, 36.004, -62.188, 37.691]
  MoveL 40 to (405.72, -210.8, 128.49) mm, rotated rx 167 ry 29.36 rz -96.45 deg; joints [118.806, 30.822, -40.814, 36.49, -60.964, 36.669]
  MoveL 41 to (403.92, -210.8, 115.73) mm, rotated rx 167 ry 29.36 rz -96.45 deg; joints [118.726, 31.984, -42.188, 36.982, -59.827, 35.779]
  MoveL 42 to (402.27, -210.8, 109.21) mm, rotated rx 167 ry 29.36 rz -96.45 deg; joints [118.653, 32.657, -42.835, 37.236, -59.279, 35.376]
  Establecer velocidad (1000.0 mm/s)
  MoveL 43 to (402.27, -210.8, 109.21) mm, rotated rx 167 ry 29.36 rz -96.45 deg; joints [118.653, 32.657, -42.835, 37.236, -59.279, 35.376]
  MoveL 44 to (421.88, -210.8, 207.27) mm, rotated rx 167 ry 29.36 rz -96.45 deg; joints [119.547, 23.84, -32.146, 33.91, -68.396, 41.654]

--- program arriderch (robot Fanuc LR Mate 200iD/7L) ---
  Suave(1)
  Establecer velocidad (1000.0 mm/s)
  Est. Ref.: RobotiQ 2F-140 Gripper (Mechanism) Base
  Est. herr: Tool 1
  Mostrar Tool 1
  MoveJ 1 to (186.94, 3.36, 269.46) mm, rotated rx 168.69 ry 0 rz -89.99 deg; joints [86.543, 38.392, -10.02, -0.729, -68.693, 93.655]
  MoveL 2 to (186.94, 3.36, 269.46) mm, rotated rx 168.69 ry 0 rz -89.99 deg; joints [86.543, 38.392, -10.02, -0.729, -68.693, 93.655]
  MoveL 3 to (167.33, 3.36, 171.4) mm, rotated rx 168.69 ry 0 rz -89.99 deg; joints [86.632, 43.937, -19.702, -0.772, -59.01, 93.7]
  MoveL 4 to (167.33, 3.36, 171.4) mm, rotated rx 168.69 ry 0 rz -89.99 deg; joints [86.632, 43.937, -19.702, -0.772, -59.01, 93.7]
  Establecer velocidad (50.0 mm/s)
  MoveL 5 to (167.33, 3.36, 181.14) mm, rotated rx 168.69 ry 0 rz -89.99 deg; joints [86.632, 43.576, -18.606, -0.764, -60.107, 93.683]
  MoveL 6 to (167.33, 3.36, 186.01) mm, rotated rx 168.69 ry 0 rz -89.99 deg; joints [86.632, 43.404, -18.052, -0.759, -60.661, 93.675]
  MoveL 7 to (167.36, 3.36, 187.22) mm, rotated rx 168.69 ry 0 rz -89.99 deg; joints [86.632, 43.357, -17.917, -0.758, -60.796, 93.673]
  MoveL 8 to (167.73, 3.36, 188.38) mm, rotated rx 168.69 ry 0 rz -89.99 deg; joints [86.63, 43.264, -17.823, -0.758, -60.889, 93.673]
  MoveL 9 to (169.47, 3.36, 190.03) mm, rotated rx 168.69 ry 0 rz -89.99 deg; joints [86.623, 42.953, -17.82, -0.76, -60.892, 93.682]
  MoveL 10 to (171.13, 3.36, 190.51) mm, rotated rx 168.69 ry 0 rz -89.99 deg; joints [86.615, 42.695, -17.942, -0.762, -60.77, 93.692]
  MoveL 11 to (172.82, 3.36, 190.92) mm, rotated rx 168.69 ry 0 rz -89.99 deg; joints [86.608, 42.436, -18.073, -0.765, -60.64, 93.702]
  MoveL 12 to (175.47, 3.36, 191.55) mm, rotated rx 168.69 ry 0 rz -89.99 deg; joints [86.596, 42.031, -18.276, -0.769, -60.436, 93.718]
  MoveL 13 to (180.22, 3.36, 192.63) mm, rotated rx 168.69 ry 0 rz -89.99 deg; joints [86.574, 41.314, -18.637, -0.777, -60.076, 93.747]
  MoveL 14 to (188.73, 3.36, 194.4) mm, rotated rx 168.69 ry 0 rz -89.99 deg; joints [86.535, 40.052, -19.275, -0.791, -59.439, 93.8]
  MoveL 15 to (210.58, 3.36, 198) mm, rotated rx 168.69 ry 0 rz -89.99 deg; joints [86.43, 36.939, -20.865, -0.829, -57.85, 93.942]
  MoveL 16 to (220.25, 3.36, 199.17) mm, rotated rx 168.69 ry 0 rz -89.99 deg; joints [86.382, 35.611, -21.555, -0.846, -57.161, 94.007]
  MoveL 17 to (224.51, 3.36, 199.6) mm, rotated rx 168.69 ry 0 rz -89.99 deg; joints [86.36, 35.036, -21.857, -0.854, -56.859, 94.037]
  MoveL 18 to (226.19, 3.36, 199.75) mm, rotated rx 168.69 ry 0 rz -89.99 deg; joints [86.351, 34.811, -21.976, -0.857, -56.74, 94.048]
  MoveL 19 to (227.87, 3.36, 199.91) mm, rotated rx 168.69 ry 0 rz -89.99 deg; joints [86.343, 34.586, -22.093, -0.861, -56.623, 94.06]
  MoveL 20 to (227.87, 3.36, 199.91) mm, rotated rx 168.69 ry 0 rz -89.99 deg; joints [86.343, 34.586, -22.093, -0.861, -56.623, 94.06]
  MoveL 21 to (240.32, 3.36, 201.51) mm, rotated rx 168.69 ry 0 rz -89.99 deg; joints [86.277, 32.916, -22.88, -0.884, -55.837, 94.148]
  MoveL 22 to (252.59, 3.36, 204.14) mm, rotated rx 168.69 ry 0 rz -89.99 deg; joints [86.21, 31.248, -23.478, -0.907, -55.24, 94.234]
  MoveL 23 to (264.62, 3.36, 207.79) mm, rotated rx 168.69 ry 0 rz -89.99 deg; joints [86.141, 29.582, -23.886, -0.927, -54.834, 94.318]
  MoveL 24 to (276.3, 3.36, 212.42) mm, rotated rx 168.69 ry 0 rz -89.99 deg; joints [86.072, 27.928, -24.099, -0.946, -54.621, 94.399]
  MoveL 25 to (290.54, 3.36, 219.68) mm, rotated rx 168.69 ry 0 rz -89.99 deg; joints [85.985, 25.851, -24.092, -0.967, -54.63, 94.497]
  MoveL 26 to (303.95, 3.36, 228.4) mm, rotated rx 168.69 ry 0 rz -89.99 deg; joints [85.9, 23.823, -23.778, -0.984, -54.945, 94.586]
  MoveL 27 to (316.37, 3.36, 238.48) mm, rotated rx 168.69 ry 0 rz -89.99 deg; joints [85.817, 21.869, -23.167, -0.996, -55.557, 94.666]
  MoveL 28 to (327.66, 3.36, 249.8) mm, rotated rx 168.69 ry 0 rz -89.99 deg; joints [85.739, 20.017, -22.276, -1.004, -56.45, 94.734]
  Establecer velocidad (1000.0 mm/s)
  MoveL 29 to (327.66, 3.36, 249.8) mm, rotated rx 168.69 ry 0 rz -89.99 deg; joints [85.739, 20.017, -22.276, -1.004, -56.45, 94.734]
  MoveL 30 to (347.27, 3.36, 347.86) mm, rotated rx 168.69 ry 0 rz -89.99 deg; joints [85.595, 14.945, -10.272, -0.93, -68.454, 94.661]
  Establecer velocidad (1000.0 mm/s)
  MoveL 31 to (428.25, 3.36, 347.86) mm, rotated rx 168.69 ry 0 rz -89.99 deg; joints [84.887, 4.47, -12.125, -1.093, -66.613, 95.448]
  MoveL 32 to (408.64, 3.36, 249.8) mm, rotated rx 168.69 ry 0 rz -89.99 deg; joints [85.079, 10.038, -25.128, -1.2, -53.609, 95.537]
  MoveL 33 to (408.64, 3.36, 249.8) mm, rotated rx 168.69 ry 0 rz -89.99 deg; joints [85.079, 10.038, -25.128, -1.2, -53.609, 95.537]
  Establecer velocidad (50.0 mm/s)
  MoveL 34 to (410.47, 3.36, 239.28) mm, rotated rx 168.69 ry 0 rz -89.99 deg; joints [85.062, 10.316, -26.607, -1.228, -52.132, 95.596]
  MoveL 35 to (412.52, 3.36, 228.8) mm, rotated rx 168.69 ry 0 rz -89.99 deg; joints [85.043, 10.601, -28.091, -1.258, -50.648, 95.659]
  MoveL 36 to (414.66, 3.36, 218.34) mm, rotated rx 168.69 ry 0 rz -89.99 deg; joints [85.022, 10.911, -29.583, -1.291, -49.157, 95.726]
  MoveL 37 to (415.77, 3.36, 208.21) mm, rotated rx 168.69 ry 0 rz -89.99 deg; joints [85.012, 11.363, -31.008, -1.323, -47.733, 95.782]
  MoveL 38 to (415.74, 3.36, 198.04) mm, rotated rx 168.69 ry 0 rz -89.99 deg; joints [85.012, 11.989, -32.411, -1.353, -46.33, 95.826]
  MoveL 39 to (414.57, 3.36, 188) mm, rotated rx 168.69 ry 0 rz -89.99 deg; joints [85.023, 12.773, -33.761, -1.382, -44.98, 95.858]
  MoveL 40 to (412.27, 3.36, 178.13) mm, rotated rx 168.69 ry 0 rz -89.99 deg; joints [85.046, 13.706, -35.048, -1.408, -43.693, 95.877]
  Establecer velocidad (1000.0 mm/s)
  MoveL 41 to (412.27, 3.36, 178.13) mm, rotated rx 168.69 ry 0 rz -89.99 deg; joints [85.046, 13.706, -35.048, -1.408, -43.693, 95.877]
  MoveL 42 to (431.88, 3.36, 276.19) mm, rotated rx 168.69 ry 0 rz -89.99 deg; joints [84.851, 6.006, -21.959, -1.208, -56.783, 95.712]

--- program arridergr (robot Fanuc LR Mate 200iD/7L) ---
  Suave(1)
  Establecer velocidad (1000.0 mm/s)
  Est. Ref.: RobotiQ 2F-140 Gripper (Mechanism) Base
  Est. herr: Tool 1
  Mostrar Tool 1
  MoveJ 1 to (354.51, 180.04, 363.6) mm, rotated rx 169.92 ry -37.62 rz -129.36 deg; joints [69.224, 31.795, -5.821, -34.789, -64.231, 77.863]
  MoveL 2 to (354.51, 180.04, 363.6) mm, rotated rx 169.92 ry -37.62 rz -129.36 deg; joints [69.224, 31.795, -5.821, -34.789, -64.231, 77.863]
  MoveL 3 to (334.9, 180.04, 265.55) mm, rotated rx 169.92 ry -37.62 rz -129.36 deg; joints [69.776, 36.105, -16.726, -38.457, -55.142, 84.888]
  MoveL 4 to (334.9, 180.04, 265.55) mm, rotated rx 169.92 ry -37.62 rz -129.36 deg; joints [69.776, 36.105, -16.726, -38.457, -55.142, 84.888]
  Establecer velocidad (50.0 mm/s)
  MoveL 5 to (332.39, 180.04, 265.31) mm, rotated rx 169.92 ry -37.62 rz -129.36 deg; joints [69.845, 36.442, -16.546, -38.363, -55.242, 84.689]
  MoveL 6 to (329.87, 180.04, 265.08) mm, rotated rx 169.92 ry -37.62 rz -129.36 deg; joints [69.913, 36.781, -16.362, -38.268, -55.345, 84.488]
  MoveL 7 to (323.48, 180.04, 264.44) mm, rotated rx 169.92 ry -37.62 rz -129.36 deg; joints [70.085, 37.652, -15.891, -38.026, -55.614, 83.977]
  MoveL 8 to (308.97, 180.04, 262.69) mm, rotated rx 169.92 ry -37.62 rz -129.36 deg; joints [70.464, 39.681, -14.786, -37.474, -56.263, 82.812]
  MoveL 9 to (276.21, 180.04, 257.29) mm, rotated rx 169.92 ry -37.62 rz -129.36 deg; joints [71.272, 44.587, -12.054, -36.196, -57.98, 80.113]
  MoveL 10 to (263.44, 180.04, 254.63) mm, rotated rx 169.92 ry -37.62 rz -129.36 deg; joints [71.57, 46.651, -10.867, -35.681, -58.77, 79.017]
  MoveL 11 to (256.31, 180.04, 253.01) mm, rotated rx 169.92 ry -37.62 rz -129.36 deg; joints [71.732, 47.849, -10.165, -35.387, -59.248, 78.39]
  MoveL 12 to (252.33, 180.04, 252.06) mm, rotated rx 169.92 ry -37.62 rz -129.36 deg; joints [71.821, 48.535, -9.759, -35.221, -59.529, 78.034]
  MoveL 13 to (249.8, 180.04, 251.45) mm, rotated rx 169.92 ry -37.62 rz -129.36 deg; joints [71.877, 48.977, -9.495, -35.115, -59.713, 77.805]
  MoveL 14 to (247.31, 180.04, 250.74) mm, rotated rx 169.92 ry -37.62 rz -129.36 deg; joints [71.933, 49.42, -9.241, -35.013, -59.889, 77.584]
  MoveL 15 to (244.7, 180.04, 248.26) mm, rotated rx 169.92 ry -37.62 rz -129.36 deg; joints [71.99, 49.913, -9.185, -34.977, -59.902, 77.494]
  MoveL 16 to (244.15, 180.04, 246.52) mm, rotated rx 169.92 ry -37.62 rz -129.36 deg; joints [72.002, 50.035, -9.325, -35.02, -59.781, 77.575]
  MoveL 17 to (244.1, 180.04, 244.7) mm, rotated rx 169.92 ry -37.62 rz -129.36 deg; joints [72.003, 50.071, -9.544, -35.093, -59.601, 77.72]
  MoveL 18 to (244.1, 180.04, 237.4) mm, rotated rx 169.92 ry -37.62 rz -129.36 deg; joints [72.003, 50.194, -10.442, -35.401, -58.868, 78.323]
  MoveL 19 to (244.1, 180.04, 222.79) mm, rotated rx 169.92 ry -37.62 rz -129.36 deg; joints [72.003, 50.494, -12.197, -36.038, -57.443, 79.529]
  Establecer velocidad (1000.0 mm/s)
  MoveL 20 to (244.1, 180.04, 222.79) mm, rotated rx 169.92 ry -37.62 rz -129.36 deg; joints [72.003, 50.494, -12.197, -36.038, -57.443, 79.529]
  MoveL 21 to (263.71, 180.04, 320.85) mm, rotated rx 169.92 ry -37.62 rz -129.36 deg; joints [71.563, 46.233, -2.168, -33.105, -65.958, 73.48]
  Establecer velocidad (1000.0 mm/s)
  MoveL 22 to (354.51, 180.04, 363.6) mm, rotated rx 169.92 ry -37.62 rz -129.36 deg; joints [69.224, 31.795, -5.821, -34.789, -64.231, 77.863]
  MoveL 23 to (334.9, 180.04, 265.55) mm, rotated rx 169.92 ry -37.62 rz -129.36 deg; joints [69.776, 36.105, -16.726, -38.457, -55.142, 84.888]
  MoveL 24 to (334.9, 180.04, 265.55) mm, rotated rx 169.92 ry -37.62 rz -129.36 deg; joints [69.776, 36.105, -16.726, -38.457, -55.142, 84.888]
  Establecer velocidad (50.0 mm/s)
  MoveL 25 to (353.58, 180.04, 267.96) mm, rotated rx 169.92 ry -37.62 rz -129.36 deg; joints [69.251, 33.627, -17.905, -39.097, -54.536, 86.27]
  MoveL 26 to (371.98, 180.04, 271.9) mm, rotated rx 169.92 ry -37.62 rz -129.36 deg; joints [68.707, 31.201, -18.75, -39.595, -54.211, 87.419]
  MoveL 27 to (390.03, 180.04, 277.37) mm, rotated rx 169.92 ry -37.62 rz -129.36 deg; joints [68.147, 28.818, -19.267, -39.945, -54.152, 88.329]
  MoveL 28 to (407.55, 180.04, 284.31) mm, rotated rx 169.92 ry -37.62 rz -129.36 deg; joints [67.576, 26.484, -19.46, -40.143, -54.351, 88.991]
  MoveL 29 to (428.92, 180.04, 295.2) mm, rotated rx 169.92 ry -37.62 rz -129.36 deg; joints [66.84, 23.596, -19.248, -40.178, -54.961, 89.474]
  MoveL 30 to (449.03, 180.04, 308.29) mm, rotated rx 169.92 ry -37.62 rz -129.36 deg; joints [66.104, 20.824, -18.541, -39.993, -55.949, 89.568]
  MoveL 31 to (467.65, 180.04, 323.41) mm, rotated rx 169.92 ry -37.62 rz -129.36 deg; joints [65.382, 18.205, -17.368, -39.623, -57.29, 89.3]
  MoveL 32 to (484.59, 180.04, 340.39) mm, rotated rx 169.92 ry -37.62 rz -129.36 deg; joints [64.69, 15.786, -15.764, -39.112, -58.952, 88.707]
  Establecer velocidad (1000.0 mm/s)
  MoveL 33 to (484.59, 180.04, 340.39) mm, rotated rx 169.92 ry -37.62 rz -129.36 deg; joints [64.69, 15.786, -15.764, -39.112, -58.952, 88.707]
  MoveL 34 to (504.2, 180.04, 438.45) mm, rotated rx 169.92 ry -37.62 rz -129.36 deg; joints [63.84, 12.395, -3.227, -35.602, -69.443, 81.008]
  Establecer velocidad (1000.0 mm/s)
  MoveL 35 to (625.68, 180.04, 438.45) mm, rotated rx 169.92 ry -37.62 rz -129.36 deg; joints [57.154, -1.514, -4.601, -37.291, -72.306, 87.55]
  MoveL 36 to (606.07, 180.04, 340.39) mm, rotated rx 169.92 ry -37.62 rz -129.36 deg; joints [58.434, 2.112, -18.03, -40.784, -61.063, 95.684]
  MoveL 37 to (606.07, 180.04, 340.39) mm, rotated rx 169.92 ry -37.62 rz -129.36 deg; joints [58.434, 2.112, -18.03, -40.784, -61.063, 95.684]
  Establecer velocidad (50.0 mm/s)
  MoveL 38 to (608.8, 180.04, 324.61) mm, rotated rx 169.92 ry -37.62 rz -129.36 deg; joints [58.261, 2.333, -20.235, -41.626, -59.511, 97.499]
  MoveL 39 to (611.88, 180.04, 308.89) mm, rotated rx 169.92 ry -37.62 rz -129.36 deg; joints [58.065, 2.599, -22.453, -42.539, -57.988, 99.396]
  MoveL 40 to (615.09, 180.04, 293.2) mm, rotated rx 169.92 ry -37.62 rz -129.36 deg; joints [57.857, 2.935, -24.689, -43.528, -56.483, 101.375]
  MoveL 41 to (616.76, 180.04, 278) mm, rotated rx 169.92 ry -37.62 rz -129.36 deg; joints [57.748, 3.5, -26.866, -44.56, -54.985, 103.292]
  MoveL 42 to (616.71, 180.04, 262.74) mm, rotated rx 169.92 ry -37.62 rz -129.36 deg; joints [57.751, 4.334, -29.059, -45.68, -53.436, 105.205]
  MoveL 43 to (614.96, 180.04, 247.69) mm, rotated rx 169.92 ry -37.62 rz -129.36 deg; joints [57.866, 5.417, -31.217, -46.876, -51.873, 107.081]
  MoveL 44 to (611.51, 180.04, 232.89) mm, rotated rx 169.92 ry -37.62 rz -129.36 deg; joints [58.089, 6.736, -33.322, -48.145, -50.312, 108.912]
  Establecer velocidad (1000.0 mm/s)
  MoveL 45 to (611.51, 180.04, 232.89) mm, rotated rx 169.92 ry -37.62 rz -129.36 deg; joints [58.089, 6.736, -33.322, -48.145, -50.312, 108.912]
  MoveL 46 to (631.12, 180.04, 330.95) mm, rotated rx 169.92 ry -37.62 rz -129.36 deg; joints [56.784, -0.329, -19.394, -41.401, -61.062, 98.054]

--- program arriizqgr (robot Fanuc LR Mate 200iD/7L) ---
  Suave(1)
  Establecer velocidad (1000.0 mm/s)
  Est. Ref.: RobotiQ 2F-140 Gripper (Mechanism) Base
  Est. herr: Tool 1
  Mostrar Tool 1
  MoveJ 1 to (331.85, -146.21, 293.73) mm, rotated rx 168.69 ry 0 rz -89.99 deg; joints [96.493, 43.21, -0.704, 1.297, -78.06, 83.364]
  MoveL 2 to (331.85, -146.21, 293.73) mm, rotated rx 168.69 ry 0 rz -89.99 deg; joints [96.493, 43.21, -0.704, 1.297, -78.06, 83.364]
  MoveL 3 to (312.23, -146.21, 195.67) mm, rotated rx 168.69 ry 0 rz -89.99 deg; joints [96.332, 47.1, -11.172, 1.339, -67.591, 83.279]
  MoveL 4 to (312.23, -146.21, 195.67) mm, rotated rx 168.69 ry 0 rz -89.99 deg; joints [96.332, 47.1, -11.172, 1.339, -67.591, 83.279]
  Establecer velocidad (50.0 mm/s)
  MoveL 5 to (300.57, -146.21, 194.29) mm, rotated rx 168.69 ry 0 rz -89.99 deg; joints [96.24, 49.161, -9.752, 1.306, -69.009, 83.412]
  MoveL 6 to (288.89, -146.21, 192.65) mm, rotated rx 168.69 ry 0 rz -89.99 deg; joints [96.151, 51.354, -8.209, 1.275, -70.55, 83.543]
  MoveL 7 to (275.98, -146.21, 190.56) mm, rotated rx 168.69 ry 0 rz -89.99 deg; joints [96.055, 53.982, -6.311, 1.241, -72.445, 83.687]
  MoveL 8 to (261.39, -146.21, 187.81) mm, rotated rx 168.69 ry 0 rz -89.99 deg; joints [95.95, 57.308, -3.818, 1.204, -74.935, 83.852]
  MoveL 9 to (248.89, -146.21, 185.14) mm, rotated rx 168.69 ry 0 rz -89.99 deg; joints [95.863, 60.641, -1.198, 1.173, -77.553, 83.997]
  MoveL 10 to (242.98, -146.21, 183.77) mm, rotated rx 168.69 ry 0 rz -89.99 deg; joints [95.823, 62.478, 0.307, 1.159, -79.057, 84.069]
  MoveL 11 to (237.72, -146.21, 182.49) mm, rotated rx 168.69 ry 0 rz -89.99 deg; joints [95.787, 64.343, 1.883, 1.146, -80.632, 84.138]
  MoveL 12 to (235.51, -146.21, 181.85) mm, rotated rx 168.69 ry 0 rz -89.99 deg; joints [95.773, 65.218, 2.629, 1.141, -81.377, 84.168]
  MoveL 13 to (234.09, -146.21, 180.92) mm, rotated rx 168.69 ry 0 rz -89.99 deg; joints [95.763, 65.792, 3.051, 1.138, -81.799, 84.186]
  MoveL 14 to (232.88, -146.21, 179.35) mm, rotated rx 168.69 ry 0 rz -89.99 deg; joints [95.755, 66.25, 3.276, 1.136, -82.024, 84.198]
  MoveL 15 to (232.37, -146.21, 177.84) mm, rotated rx 168.69 ry 0 rz -89.99 deg; joints [95.752, 66.393, 3.207, 1.135, -81.955, 84.2]
  MoveL 16 to (232.28, -146.21, 176.01) mm, rotated rx 168.69 ry 0 rz -89.99 deg; joints [95.751, 66.317, 2.883, 1.136, -81.631, 84.194]
  MoveL 17 to (232.28, -146.21, 173.53) mm, rotated rx 168.69 ry 0 rz -89.99 deg; joints [95.751, 66.169, 2.399, 1.138, -81.147, 84.185]
  MoveL 18 to (232.28, -146.21, 169.12) mm, rotated rx 168.69 ry 0 rz -89.99 deg; joints [95.751, 65.941, 1.577, 1.14, -80.325, 84.168]
  MoveL 19 to (232.28, -146.21, 164.01) mm, rotated rx 168.69 ry 0 rz -89.99 deg; joints [95.751, 65.723, 0.67, 1.144, -79.418, 84.15]
  MoveL 20 to (232.28, -146.21, 158.89) mm, rotated rx 168.69 ry 0 rz -89.99 deg; joints [95.751, 65.548, -0.197, 1.147, -78.552, 84.132]
  MoveL 21 to (232.28, -146.21, 153.63) mm, rotated rx 168.69 ry 0 rz -89.99 deg; joints [95.751, 65.406, -1.048, 1.151, -77.7, 84.114]
  Establecer velocidad (1000.0 mm/s)
  MoveL 22 to (232.28, -146.21, 153.63) mm, rotated rx 168.69 ry 0 rz -89.99 deg; joints [95.751, 65.406, -1.048, 1.151, -77.7, 84.114]
  MoveL 23 to (251.89, -146.21, 251.69) mm, rotated rx 168.69 ry 0 rz -89.99 deg; joints [95.883, 64.283, 11.433, 1.15, -90.182, 84.234]
  Establecer velocidad (1000.0 mm/s)
  MoveL 24 to (343.61, -146.21, 294.87) mm, rotated rx 168.69 ry 0 rz -89.99 deg; joints [96.593, 41.055, -2.06, 1.324, -76.707, 83.229]
  MoveL 25 to (323.99, -146.21, 196.81) mm, rotated rx 168.69 ry 0 rz -89.99 deg; joints [96.428, 45.132, -12.508, 1.372, -66.258, 83.143]
  MoveL 26 to (323.99, -146.21, 196.81) mm, rotated rx 168.69 ry 0 rz -89.99 deg; joints [96.428, 45.132, -12.508, 1.372, -66.258, 83.143]
  Establecer velocidad (50.0 mm/s)
  MoveL 27 to (346.2, -146.21, 199.83) mm, rotated rx 168.69 ry 0 rz -89.99 deg; joints [96.616, 41.612, -14.646, 1.437, -64.125, 82.884]
  MoveL 28 to (370.59, -146.21, 205.77) mm, rotated rx 168.69 ry 0 rz -89.99 deg; joints [96.836, 37.903, -16.345, 1.507, -62.432, 82.598]
  MoveL 29 to (394.18, -146.21, 214.34) mm, rotated rx 168.69 ry 0 rz -89.99 deg; joints [97.063, 34.38, -17.371, 1.571, -61.412, 82.321]
  MoveL 30 to (416.7, -146.21, 225.43) mm, rotated rx 168.69 ry 0 rz -89.99 deg; joints [97.294, 31.022, -17.767, 1.629, -61.023, 82.057]
  MoveL 31 to (437.87, -146.21, 238.92) mm, rotated rx 168.69 ry 0 rz -89.99 deg; joints [97.526, 27.833, -17.563, 1.677, -61.233, 81.812]
  MoveL 32 to (457.44, -146.21, 254.64) mm, rotated rx 168.69 ry 0 rz -89.99 deg; joints [97.753, 24.838, -16.795, 1.715, -62.007, 81.591]
  MoveL 33 to (475.18, -146.21, 272.4) mm, rotated rx 168.69 ry 0 rz -89.99 deg; joints [97.971, 22.077, -15.502, 1.742, -63.306, 81.399]
  Establecer velocidad (1000.0 mm/s)
  MoveL 34 to (475.18, -146.21, 272.4) mm, rotated rx 168.69 ry 0 rz -89.99 deg; joints [97.971, 22.077, -15.502, 1.742, -63.306, 81.399]
  MoveL 35 to (494.79, -146.21, 370.46) mm, rotated rx 168.69 ry 0 rz -89.99 deg; joints [98.226, 18.374, -3.445, 1.66, -75.365, 81.512]
  Establecer velocidad (1000.0 mm/s)
  MoveL 36 to (625.33, -146.21, 329.23) mm, rotated rx 168.69 ry 0 rz -89.99 deg; joints [100.453, 1.718, -12.093, 2.216, -66.796, 78.872]
  MoveL 37 to (605.72, -146.21, 231.17) mm, rotated rx 168.69 ry 0 rz -89.99 deg; joints [100.046, 7.319, -25.385, 2.437, -53.499, 78.695]
  MoveL 38 to (605.72, -146.21, 231.17) mm, rotated rx 168.69 ry 0 rz -89.99 deg; joints [100.046, 7.319, -25.385, 2.437, -53.499, 78.695]
  Establecer velocidad (50.0 mm/s)
  MoveL 39 to (608.5, -146.21, 212.05) mm, rotated rx 168.69 ry 0 rz -89.99 deg; joints [100.102, 7.939, -28.096, 2.542, -50.794, 78.482]
  MoveL 40 to (608.54, -146.21, 192.73) mm, rotated rx 168.69 ry 0 rz -89.99 deg; joints [100.103, 9.028, -30.802, 2.647, -48.09, 78.32]
  MoveL 41 to (605.85, -146.21, 173.61) mm, rotated rx 168.69 ry 0 rz -89.99 deg; joints [100.049, 10.551, -33.426, 2.749, -45.467, 78.213]
  MoveL 42 to (603.37, -146.21, 163.83) mm, rotated rx 168.69 ry 0 rz -89.99 deg; joints [100, 11.499, -34.733, 2.799, -44.159, 78.181]
  Establecer velocidad (1000.0 mm/s)
  MoveL 43 to (603.37, -146.21, 163.83) mm, rotated rx 168.69 ry 0 rz -89.99 deg; joints [100, 11.499, -34.733, 2.799, -44.159, 78.181]
  MoveL 44 to (622.98, -146.21, 261.88) mm, rotated rx 168.69 ry 0 rz -89.99 deg; joints [100.403, 3.857, -21.35, 2.403, -57.544, 78.504]

